ACTION act_Status:
IF TRUE 
AND fbPis.m_CheckByRecipe(stPis:=stPis_TankA, 			req:=E_Piston_Recipe_State.Release)	
//AND fbPis.m_CheckByRecipe(stPis:=stPis_TankA_Pipe, 		req:=E_Piston_Recipe_State.Release)	
AND fbPis.m_CheckByRecipe(stPis:=stPis_TankB, 			req:=E_Piston_Recipe_State.Release)
//AND fbPis.m_CheckByRecipe(stPis:=stPis_TankB_Pipe, 		req:=E_Piston_Recipe_State.Release)
AND fbPis.m_CheckByRecipe(stPis:=stPis_Drain, 			req:=E_Piston_Recipe_State.Release)
AND fbPis.m_CheckByRecipe(stPis:=stPis_CIP, 			req:=E_Piston_Recipe_State.Release)
THEN;
	eStatus:=E_Line_Target.eClose;
ELSIF TRUE 
AND fbPis.m_CheckByRecipe(stPis:=stPis_TankA, 			req:=E_Piston_Recipe_State.Act)		
AND fbPis.m_CheckByRecipe(stPis:=stPis_TankA_Pipe, 		req:=E_Piston_Recipe_State.Release)	
AND fbPis.m_CheckByRecipe(stPis:=stPis_TankB, 			req:=E_Piston_Recipe_State.Release)
//AND fbPis.m_CheckByRecipe(stPis:=stPis_TankB_Pipe, 		req:=E_Piston_Recipe_State.Release)
AND fbPis.m_CheckByRecipe(stPis:=stPis_Drain, 			req:=E_Piston_Recipe_State.Release)
AND fbPis.m_CheckByRecipe(stPis:=stPis_CIP, 			req:=E_Piston_Recipe_State.Release)
THEN;
	eStatus:=E_Line_Target.eTank_A;
ELSIF TRUE 
AND fbPis.m_CheckByRecipe(stPis:=stPis_TankA, 			req:=E_Piston_Recipe_State.Release)		
//AND fbPis.m_CheckByRecipe(stPis:=stPis_TankA_Pipe, 		req:=E_Piston_Recipe_State.Release)	
AND fbPis.m_CheckByRecipe(stPis:=stPis_TankB, 			req:=E_Piston_Recipe_State.Act)
AND fbPis.m_CheckByRecipe(stPis:=stPis_TankB_Pipe, 		req:=E_Piston_Recipe_State.Release)
AND fbPis.m_CheckByRecipe(stPis:=stPis_Drain, 			req:=E_Piston_Recipe_State.Release)
AND fbPis.m_CheckByRecipe(stPis:=stPis_CIP, 			req:=E_Piston_Recipe_State.Release)
THEN;
	eStatus:=E_Line_Target.eTank_B;
ELSIF TRUE 
AND fbPis.m_CheckByRecipe(stPis:=stPis_TankA, 			req:=E_Piston_Recipe_State.Release)		
//AND fbPis.m_CheckByRecipe(stPis:=stPis_TankA_Pipe, 		req:=E_Piston_Recipe_State.Release)	
AND fbPis.m_CheckByRecipe(stPis:=stPis_TankB, 			req:=E_Piston_Recipe_State.Release)
//AND fbPis.m_CheckByRecipe(stPis:=stPis_TankB_Pipe, 		req:=E_Piston_Recipe_State.Release)
AND fbPis.m_CheckByRecipe(stPis:=stPis_Drain, 			req:=E_Piston_Recipe_State.Act)
AND fbPis.m_CheckByRecipe(stPis:=stPis_CIP, 			req:=E_Piston_Recipe_State.Act)
THEN;
	eStatus:=E_Line_Target.eCIP;
ELSIF TRUE 
AND fbPis.m_CheckByRecipe(stPis:=stPis_TankA, 			req:=E_Piston_Recipe_State.Release)		
//AND fbPis.m_CheckByRecipe(stPis:=stPis_TankA_Pipe, 		req:=E_Piston_Recipe_State.Release)	
AND fbPis.m_CheckByRecipe(stPis:=stPis_TankB, 			req:=E_Piston_Recipe_State.Release)
//AND fbPis.m_CheckByRecipe(stPis:=stPis_TankB_Pipe, 		req:=E_Piston_Recipe_State.Release)
AND fbPis.m_CheckByRecipe(stPis:=stPis_Drain, 			req:=E_Piston_Recipe_State.Act)
AND fbPis.m_CheckByRecipe(stPis:=stPis_CIP, 			req:=E_Piston_Recipe_State.Release)
THEN;
	eStatus:=E_Line_Target.eDrain;
ELSE;
	eStatus:=E_Line_Target.eNone;
END_IF
END_ACTION

METHOD m_CheckStatus : BOOL
VAR_INPUT
	eReqStatus		: E_Line_Target;
END_VAR
IF eStatus=eReqStatus 
AND eProcess=E_Line_Target.eNone
AND eReq=E_Line_Target.eNone
AND bReady
AND bDone
AND NOT bRun
THEN;
	m_CheckStatus:=TRUE;
END_IF
END_METHOD

METHOD m_Request_Reset : BOOL
VAR_IN_OUT
	memo: R_TRIG;
END_VAR
memo(CLK:=eReq=0);
IF TRUE 
AND memo.Q
THEN;
	SFCReset:=TRUE;
END_IF
END_METHOD

METHOD m_Run : BOOL
VAR_INPUT
	eReqProc			: E_Line_Target;
END_VAR
IF eProcess=E_Line_Target.eNone THEN;
	eProcess:=eReq:=eReqProc;
	bDone:=FALSE;
	m_Run:=TRUE;
END_IF
END_METHOD

METHOD m_Set_SFCFlags_Reference : BOOL
//Set reference to SFC flags

refSFC.SFCInit REF= SFCInit;
refSFC.SFCReset REF= SFCReset;
refSFC.SFCError REF= SFCError;
refSFC.SFCEnableLimit REF= SFCEnableLimit;
refSFC.SFCErrorStep REF= SFCErrorStep;
refSFC.SFCErrorPOU REF= SFCErrorPOU;
refSFC.SFCQuitError REF= SFCQuitError;
refSFC.SFCPause REF= SFCPause;
refSFC.SFCTrans REF= SFCTrans;
refSFC.SFCCurrentStep REF= SFCCurrentStep;
refSFC.SFCTip REF= SFCTip;
refSFC.SFCTipMode REF= SFCTipMode;

// Cycle handle for SFC
m_SFC_Handle();
END_METHOD

END_FUNCTION_BLOCK

// ---- 00 Library/02 Pump/FB_Pump.TcPOU
FUNCTION_BLOCK FB_Pump
VAR_INPUT
	Pump_ID				: E_Pump_List:=E_Pump_List.eNotSelected;
	PressureSensor_ID	: E_ASense_Name:=E_ASense_Name.eNotSelected;
END_VAR
VAR
	sID: STRING(6);

	stNidec: REFERENCE TO ST_Nidec;
	status_word: WORD;
	control_word: WORD;

	ControlWord: ControlWordStruct;
	StatusWord: StatusWordStruct;


	//request
	modeAuto	:	BOOL	:= TRUE	;//System in automatic
	bRun_Auto	:	BOOL	;
	bRun_Man	:	BOOL	;

	//nRPM_Auto	:	REAL		;//Pump RPM 
	//nRPM_Man	:	REAL		;//Pump RPM 
	//feedback
	nRPM_fdbk	:	INT	;	
	rtManual: R_TRIG;
	ton_Drive_init: TON;
	state_init: (OFF,stage1,stage2,stage3,stage4, Ready);

	bInitiated: BOOL;
	ton_RPM_feedback_lag_monitoring: TON;
	ton_Pressure_feedback_monitoring: TON;
	
	fbPressureSensor: REFERENCE TO FB_AnalogSensor;

END_VAR
VAR_OUTPUT
	DriveReady	:   BOOL;
	bRun		: 	BOOL;
	nRPM		:	REAL		;//Pump RPM 
	
END_VAR
VAR_IN_OUT
	stPump			: ST_Pump	;
	stOperation		: ST_OperationButtons;
END_VAR

stNidec REF= gIO.Nidec[Pump_ID];
sID:=TO_STRING(Pump_ID);
nRPM:=stPump.nRPM;
IF __ISVALIDREF(stNidec) THEN;
	//run
	status_word:=stNidec.StatusWord;
	stNidec.ControlWord:=control_word;
	
	control_word:=m_Map_ControlWord(cwStruct:=ControlWord);
	StatusWord:=m_Map_StatusWord(wordInput:=status_word);
	
	stNidec.targetVelocity:=DINT_TO_INT(TRUNC(stPump.nRPM));	
	nRPM_fdbk:=stNidec.actVelocity;	
	
	m_Nidec_Init();
	
	IF state_init=Ready THEN;
		DriveReady:=TRUE;
		ControlWord.EnableOperation:=bRun;
	ELSE;
		DriveReady:=FALSE;
		//bRun:=bRun_Man:=bRun_Auto:=FALSE;
		ControlWord.EnableOperation:=FALSE;
	END_IF	
	stPump.DriveReady:=DriveReady;
ELSE;
	//RETURN;
END_IF

IF modeAuto THEN;
	//bRun:=bRun_Auto;
	IF bRun_Auto AND m_CheckOper() THEN;
		bRun:=TRUE;
	ELSE;
		bRun:=FALSE;
	END_IF
	stPump.nRPM:=stPump.nRPM_Auto;
ELSE;
	//bRun:=bRun_Man;
	IF bRun_Man AND m_CheckOper() THEN;
		bRun:=TRUE;
	ELSE;
		bRun:=FALSE;
	END_IF	
	stPump.nRPM:=stPump.nRPM_Man;
END_IF

rtManual(CLK:=NOT modeAuto);
IF rtManual.Q THEN;
	bRun:=bRun_Man:=bRun_Auto;
	//stPump.nRPM:=stPump.nRPM_Man:=stPump.nRPM_Auto;
END_IF

IF stPump.nRPM>3000 THEN;
	stPump.nRPM:=3000;
END_IF

stPump.bRun_Man:=bRun_Man;
stPump.bRun_Auto:=bRun_Auto;
stPump.bRun:=bRun;

IF m_Error()<>'' THEN;
	//stOperation.bSetPause:=TRUE;
	//print error
	//fbPrintErrMessageByID(sModuleDescription:='Pump',sActErrorID:='101x000x001');	
END_IF

bInitiated:=TRUE;

METHOD m_Auto : BOOL
VAR_INPUT
	control: LREAL; // RPM
END_VAR

VAR
	RPM: INT;
END_VAR
//ST_Pump.bRun_Auto:=TRUE;
m_Auto:=TRUE;
RPM:=DINT_TO_INT(TRUNC(control));
IF RPM>3000 THEN;
	stPump.nRPM_Auto:=3000;
ELSIF RPM<200 THEN;
	stPump.nRPM_Auto:=200;
ELSE;
	stPump.nRPM_Auto:=RPM;
END_IF

bRun_Auto:=TRUE;
//need to be set up an set point so the pump could keep the needed value in automatic mode
END_METHOD

METHOD INTERNAL m_CheckOper : BOOL
VAR_INPUT
END_VAR

VAR
	sMotorTypeAgrigate_to_check: STRING(2);
END_VAR
sMotorTypeAgrigate_to_check:=TO_STRING(Pump_ID);

IF sMotorTypeAgrigate_to_check='AG' THEN;
	m_CheckOper:=TRUE;
ELSE;
	IF stOperation.iActOperation=E_OperationButtons.ePlayAll THEN;
		m_CheckOper:=TRUE;
	ELSE;
		m_CheckOper:=FALSE;
	END_IF
END_IF
END_METHOD

METHOD m_Error : STRING(11)
VAR_INPUT
	
END_VAR
VAR
	skipTemp: BOOL;
END_VAR
ton_RPM_feedback_lag_monitoring(PT:=T#10S);
IF __ISVALIDREF(stNidec) THEN;
	IF bRun
	AND ABS(stNidec.targetVelocity - nRPM_fdbk) > 10 
	THEN;
		ton_RPM_feedback_lag_monitoring.IN:=TRUE;
	ELSE;
		ton_RPM_feedback_lag_monitoring.IN:=FALSE;
	END_IF	
END_IF

CASE Pump_ID OF
	E_Pump_List.AG3001,
	E_Pump_List.AG3002,
	E_Pump_List.P3001,
	E_Pump_List.P3002:;
		skipTemp:=TRUE;
ELSE;
		skipTemp:=FALSE;
END_CASE


IF bRun AND NOT skipTemp THEN;
	IF NOT DriveReady THEN;
		m_Error:=concat(sID,'x001');
		stOperation.bSetPause:=TRUE;
		RETURN;
	END_IF	

	IF ton_RPM_feedback_lag_monitoring.Q THEN;
		m_Error:=concat(sID,'x002');
		RETURN;
	END_IF
END_IF

IF NOT DriveReady AND NOT skipTemp THEN;
	m_Error:=concat(sID,'x003');
	//stOperation.bSetPause:=TRUE;
	RETURN;
END_IF


IF 	PressureSensor_ID <> E_ASense_Name.eNotSelected THEN;
	fbPressureSensor REF= fbAnalogSensor[PressureSensor_ID];
	IF __ISVALIDREF(fbPressureSensor) THEN;	
		ton_Pressure_feedback_monitoring(PT:=T#30S);
		IF bRun AND ( fbPressureSensor.bHH_Alarm 
					OR fbPressureSensor.bHH_Warning
					OR fbPressureSensor.bLL_Warning 
					OR fbPressureSensor.bLL_Alarm) 
		THEN;
			ton_Pressure_feedback_monitoring.IN:=TRUE;
		ELSE;
			ton_Pressure_feedback_monitoring.IN:=FALSE;
		END_IF	
		
		IF fbPressureSensor.bHH_Alarm AND ton_Pressure_feedback_monitoring.Q THEN;
			m_Error:=concat(sID,'x004');
			stOperation.bSetPause:=TRUE;
			RETURN;
		END_IF
		IF fbPressureSensor.bHH_Warning AND ton_Pressure_feedback_monitoring.Q THEN;
			m_Error:=concat(sID,'x005');
			RETURN;
		END_IF
		IF fbPressureSensor.bLL_Warning AND ton_Pressure_feedback_monitoring.Q THEN;
			m_Error:=concat(sID,'x006');
			RETURN;
		END_IF
		IF fbPressureSensor.bLL_Alarm AND ton_Pressure_feedback_monitoring.Q THEN;
			m_Error:=concat(sID,'x007');
			stOperation.bSetPause:=TRUE;
			RETURN;
		END_IF		
	END_IF	
END_IF

IF NOT modeAuto THEN;
	m_Error:=concat(sID,'x008');
	//stOperation.bSetPause:=TRUE;
	RETURN;
END_IF

m_Error:='';
END_METHOD

METHOD m_Get_Speed : INT
VAR_INPUT
END_VAR
m_Get_Speed:=nRPM_fdbk;
END_METHOD

METHOD m_Map_ControlWord : WORD
VAR_INPUT
	cwStruct : ControlWordStruct;
END_VAR
VAR
    tempWord : WORD;
END_VAR


// Map each bit from the structure to the corresponding bit in the control word
tempWord := 0;
IF cwStruct.SwitchOn THEN
    tempWord := tempWord OR 1; // Bit 0
END_IF
IF cwStruct.EnableVoltage THEN
    tempWord := tempWord OR 2; // Bit 1
END_IF
IF cwStruct.QuickStop THEN
    tempWord := tempWord OR 4; // Bit 2
END_IF
IF cwStruct.EnableOperation THEN
    tempWord := tempWord OR 8; // Bit 3
END_IF
// Reserved bits (4-7) are not set
IF cwStruct.FaultReset THEN
    tempWord := tempWord OR 256; // Bit 8
END_IF
// Reserved bits (9-15) are not set

m_Map_ControlWord := tempWord;
END_METHOD

METHOD m_Map_StatusWord : StatusWordStruct
VAR_INPUT
	wordInput : WORD;
END_VAR
VAR
    swStruct : StatusWordStruct;
END_VAR


// Map each bit from the status word to the corresponding field in the structure
swStruct.ReadyToSwitchOn    := (wordInput AND 1) <> 0;         // Bit 0
swStruct.SwitchedOn         := (wordInput AND 2) <> 0;         // Bit 1
swStruct.OperationEnabled   := (wordInput AND 4) <> 0;         // Bit 2
swStruct.Fault              := (wordInput AND 8) <> 0;         // Bit 3
swStruct.VoltageEnabled     := (wordInput AND 16) <> 0;        // Bit 4
swStruct.QuickStop          := (wordInput AND 32) <> 0;        // Bit 5
swStruct.SwitchOnDisabled   := (wordInput AND 64) <> 0;        // Bit 6
swStruct.Warning            := (wordInput AND 128) <> 0;       // Bit 7
swStruct.Remote             := (wordInput AND 256) <> 0;       // Bit 8
// Reserved bits (9-15) are not set, assuming FALSE
m_Map_StatusWord := swStruct;
END_METHOD

METHOD m_Nidec_Init : BOOL
VAR_INPUT
END_VAR
IF  NOT StatusWord.VoltageEnabled 
OR StatusWord.Fault 
OR (state_init=Ready AND NOT StatusWord.ReadyToSwitchOn )
THEN;
	ControlWord.SwitchOn:=FALSE;
	ControlWord.EnableVoltage:=FALSE;
	ControlWord.QuickStop:=FALSE;
	ControlWord.EnableOperation:=FALSE;
	ton_Drive_init(IN:=FALSE);
	state_init:=OFF;
	RETURN;
END_IF


CASE state_init OF
	OFF:; 
		IF TRUE
		AND StatusWord.VoltageEnabled
		AND StatusWord.QuickStop
		AND StatusWord.SwitchOnDisabled
		THEN;
			ton_Drive_init(IN:=TRUE,PT:=T#2S);
		ELSE;
			ton_Drive_init(IN:=FALSE);RETURN;
		END_IF
		
		IF ton_Drive_init.Q THEN;
			ControlWord.EnableVoltage:=TRUE;
			ControlWord.QuickStop:=TRUE;	
			state_init:=stage1;
			ton_Drive_init(IN:=FALSE);
		END_IF	
		
	stage1:;
		IF TRUE
		AND StatusWord.VoltageEnabled
		AND StatusWord.QuickStop
		AND NOT StatusWord.SwitchOnDisabled
		THEN;
			ton_Drive_init(IN:=TRUE,PT:=T#0.5S);
		ELSE;
			ton_Drive_init(IN:=FALSE);RETURN;
		END_IF
		
		IF ton_Drive_init.Q THEN;
			ControlWord.SwitchOn:=TRUE;
			state_init:=stage2;
			ton_Drive_init(IN:=FALSE);
		END_IF	
		
	stage2:;
		IF TRUE
		AND StatusWord.SwitchedOn
		AND StatusWord.VoltageEnabled
		AND StatusWord.QuickStop
		AND NOT StatusWord.SwitchOnDisabled
		THEN;
			ton_Drive_init(IN:=TRUE,PT:=T#0.5S);
		ELSE;
			ton_Drive_init(IN:=FALSE);RETURN;
		END_IF
		
		IF ton_Drive_init.Q THEN;
			state_init:=Ready;
			ton_Drive_init(IN:=FALSE);
		END_IF	

	
	
END_CASE
END_METHOD

METHOD m_Run : BOOL
VAR_INPUT
	RPM: REAL;
END_VAR
IF NOT bInitiated THEN;
	RETURN;
END_IF
bRun_Auto:=TRUE;
stPump.nRPM_Auto:=RPM;
m_Run:=TRUE;
END_METHOD

METHOD m_Stop : BOOL
VAR_INPUT
END_VAR
bRun_Auto:=FALSE;
bRun_Man:=FALSE;
m_Stop:=TRUE;
END_METHOD

END_FUNCTION_BLOCK

// ---- 00 Library/02 Pump/02.1 Dosing Pump/FB_DosingPump.TcPOU
FUNCTION_BLOCK FB_DosingPump EXTENDS FB_SFC_Cycle
VAR_INPUT
END_VAR
VAR_OUTPUT
	valve_A			: BOOL;
	valve_B			: BOOL;
END_VAR
VAR

	action_Time		: TIME:=T#0.5S;
	startDelay		: TIME:=T#0S;
	
	reqTiks			: DINT:=5;
	actTiks			: DINT:=5;
	
	fStageVolume	: REAL:=65; 	// CC/stage
	fReqVolume		: REAL:=500.0; 	// CC
	fActVolume		: REAL; 		// CC


END_VAR

VAR PERSISTENT
	
END_VAR

act_GetReference();

act_Oper();

reqTiks:=TRUNC(fReqVolume/fStageVolume);
fActVolume:=(actTiks*fStageVolume);

ACTION _acheck_Count_active:
bStepDone:=FALSE;
IF actTiks>=reqTiks THEN;
	bStepDone:=TRUE;
END_IF
END_ACTION

ACTION _acheck_Count_entry:
actTiks:=actTiks+1;
END_ACTION

ACTION _aDone_entry:
bRun:=FALSE;
bDone:=TRUE;
END_ACTION

ACTION _aInit_act_Oper_active:
SFCReset:=FALSE;
END_ACTION

ACTION _aInit_act_Oper_exit:
valve_A:=valve_B:=bRun:=bDone:=FALSE;
END_ACTION

ACTION _aReady_exit:
actTiks:=0;
END_ACTION

ACTION _astage_A_entry:
valve_A:=TRUE;
END_ACTION

ACTION _astage_A_exit:
valve_A:=FALSE;
END_ACTION

ACTION _astage_B_entry:
valve_B:=TRUE;
END_ACTION

ACTION _astage_B_exit:
valve_B:=FALSE;
END_ACTION

ACTION act_GetReference:
m_Set_SFCFlags_Reference();
END_ACTION

ACTION act_Oper:
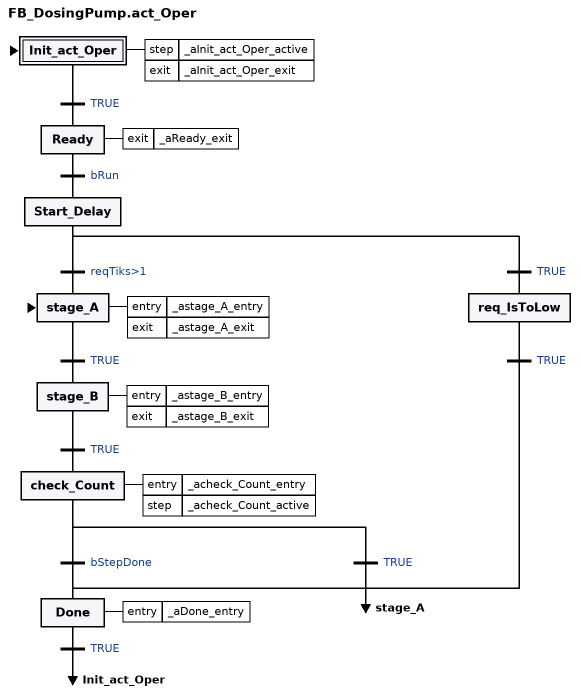
INITIAL_STEP Init_act_Oper:
    _aInit_act_Oper_active(N);  // step action
    _aInit_act_Oper_exit(P0);  // exit action
END_STEP
TRANSITION FROM Init_act_Oper TO Ready
    := TRUE;
END_TRANSITION
STEP Ready:
    _aReady_exit(P0);  // exit action
END_STEP
TRANSITION FROM Ready TO Start_Delay
    := bRun;
END_TRANSITION
STEP Start_Delay:  // min time startDelay
END_STEP
TRANSITION FROM Start_Delay TO stage_A
    := reqTiks>1;
END_TRANSITION
STEP stage_A:  // min time action_Time
    _astage_A_entry(P1);  // entry action
    _astage_A_exit(P0);  // exit action
END_STEP
TRANSITION FROM stage_A TO stage_B
    := TRUE;
END_TRANSITION
STEP stage_B:  // min time action_Time
    _astage_B_entry(P1);  // entry action
    _astage_B_exit(P0);  // exit action
END_STEP
TRANSITION FROM stage_B TO check_Count
    := TRUE;
END_TRANSITION
STEP check_Count:
    _acheck_Count_entry(P1);  // entry action
    _acheck_Count_active(N);  // step action
END_STEP
TRANSITION FROM check_Count TO Done
    := bStepDone;
END_TRANSITION
TRANSITION FROM check_Count TO stage_A
    := TRUE;
END_TRANSITION
TRANSITION FROM Start_Delay TO req_IsToLow
    := TRUE;
END_TRANSITION
STEP req_IsToLow:
END_STEP
TRANSITION FROM req_IsToLow TO Done
    := TRUE;
END_TRANSITION
STEP Done:
    _aDone_entry(P1);  // entry action
END_STEP
TRANSITION FROM Done TO Init_act_Oper
    := TRUE;
END_TRANSITION
// branch label Branch0_act_Oper
// branch label Branch1_act_Oper
END_ACTION

METHOD m_RunVolume : BOOL
VAR_INPUT
	Volume	:REAL;
END_VAR
fReqVolume:=Volume;
mRun();
IF rtDone.Q THEN;
	m_RunVolume:=TRUE;	
END_IF
END_METHOD

METHOD m_Set_SFCFlags_Reference : BOOL
//Set reference to SFC flags

refSFC.SFCInit REF= SFCInit;
refSFC.SFCReset REF= SFCReset;
refSFC.SFCError REF= SFCError;
refSFC.SFCEnableLimit REF= SFCEnableLimit;
refSFC.SFCErrorStep REF= SFCErrorStep;
refSFC.SFCErrorPOU REF= SFCErrorPOU;
refSFC.SFCQuitError REF= SFCQuitError;
refSFC.SFCPause REF= SFCPause;
refSFC.SFCTrans REF= SFCTrans;
refSFC.SFCCurrentStep REF= SFCCurrentStep;
refSFC.SFCTip REF= SFCTip;
refSFC.SFCTipMode REF= SFCTipMode;

// Cycle handle for SFC
m_SFC_Handle();
END_METHOD

METHOD m_Stop : BOOL
VAR_INPUT
END_VAR
SFCReset:=TRUE;
END_METHOD

END_FUNCTION_BLOCK

// ---- 00 Library/HeatExchenger/FB_HeatExchanger.TcPOU
FUNCTION_BLOCK FB_HeatExchanger
VAR_IN_OUT
	stHeatExchanger	:	ST_HeatExchanger	;
END_VAR
VAR_INPUT
	nValveID		:	E_Pis_Name 	;	
	nAnalogValveID	:	E_Pis_Name 	;

	nProcCntrlID	:	E_ProcessControl_Name	;
END_VAR
VAR_OUTPUT
	nAlagonValveCntrOut	:	INT	;//output for analog valve opening
END_VAR
VAR
	stPis			:	REFERENCE TO ST_Piston;
	stPisAnalog		:	REFERENCE TO ST_Piston;
	
	stProcessControl		:	REFERENCE TO ST_ProcessControl	;
	fbProcessControl		: 	REFERENCE TO FB_ProcessControl	;
END_VAR

act_GetReference();
//act_AnalogOutScaling();

stProcessControl.fCtrlOutput_Min:=0;
stProcessControl.fCtrlOutput_Max:=100;
stProcessControl.fCtrlOutput_Manual;
stProcessControl.rValue_Min_To_ReleaseControl:=15; //Degrees

IF stHeatExchanger.bManual THEN;
	fbProcessControl.mRun_PID(Set_Point:=stProcessControl.fCtrlOutput_Manual , controlManual:=TRUE);
	//nAlagonValveCntrOut:=mCMD_to_Analog(fControl:=stHeatExchanger.fManualControl);
ELSE;
	IF stProcessControl.bActiveCntr AND NOT stPis.st_Open THEN
		stPis.req_Open:=TRUE;
	ELSIF NOT stProcessControl.bActiveCntr AND NOT stPis.st_Close THEN
		stPis.req_Close:=TRUE;
	END_IF
	//nAlagonValveCntrOut:=mCMD_to_Analog(fControl:=stProcessControl.fCtrlOutput);	
END_IF
nAlagonValveCntrOut:=mCMD_to_Analog(fControl:=stProcessControl.fCtrlOutput);
IF nAlagonValveCntrOut=0 AND NOT stPisAnalog.st_Close THEN;
	stPisAnalog.req_Close:=TRUE;
ELSIF nAlagonValveCntrOut<>0 AND NOT stPisAnalog.st_Open THEN;
	stPisAnalog.req_Open:=TRUE;
END_IF

ACTION act_AnalogOutScaling:
IF (stHeatExchanger.cntrlVal_Max-stHeatExchanger.cntrlVal_Min)<>0 THEN
	nAlagonValveCntrOut:=DINT_TO_INT((TRUNC((stProcessControl.fCtrlOutput*
		(stHeatExchanger.outVal_Max-stHeatExchanger.outVal_Min)/(stHeatExchanger.cntrlVal_Max-stHeatExchanger.cntrlVal_Min))+
		stHeatExchanger.outOffset)));
END_IF
END_ACTION

ACTION act_GetReference:
//On-Off walve structure
stPis REF= g_Piston.stPis[nValveID];
stPisAnalog REF= g_Piston.stPis[nAnalogValveID];

stProcessControl REF=g_ProcControl.arr_stProcCntrl[nProcCntrlID];
fbProcessControl REF=g_ProcControl.arr_fbProcCntrl[nProcCntrlID];
END_ACTION

METHOD m_Auto : BOOL
VAR_INPUT
END_VAR
END_METHOD

METHOD m_Run : BOOL
VAR_INPUT
END_VAR
END_METHOD

METHOD m_Stop : BOOL
VAR_INPUT
END_VAR
END_METHOD

METHOD mCMD_to_Analog : INT
VAR_INPUT
	fControl: LREAL;
END_VAR
IF (stHeatExchanger.cntrlVal_Max-stHeatExchanger.cntrlVal_Min)<>0 THEN
	mCMD_to_Analog:=DINT_TO_INT((TRUNC((fControl*
		(stHeatExchanger.outVal_Max-stHeatExchanger.outVal_Min)/(stHeatExchanger.cntrlVal_Max-stHeatExchanger.cntrlVal_Min))+
		stHeatExchanger.outOffset)));
ELSE;
	mCMD_to_Analog:=0;
END_IF

//nAlagonValveCntrOut
END_METHOD

END_FUNCTION_BLOCK

// ---- 03 Project/23 CIP/FB_CIP_ClientTank.TcPOU
FUNCTION_BLOCK FB_CIP_ClientTank EXTENDS FB_SFC_Cycle IMPLEMENTS ITF_FB_SFC_Cycle
VAR_INPUT	
	valTank_A				: E_Pis_Name;
	valTank_A_Sprinkler		: E_Pis_Name;
	valTank_A_Main			: E_Pis_Name;
	valTank_B				: E_Pis_Name;
	valTank_B_Sprinkler		: E_Pis_Name;	
	valTank_B_Main			: E_Pis_Name;	
	valDrain				: E_Pis_Name;
END_VAR
VAR_OUTPUT
END_VAR
VAR

	eReq				: E_CIP_ClientTank;
	eProcess			: E_CIP_ClientTank;
	eStatus				: E_CIP_ClientTank;
	
	fbPis					: FB_Piston;
	stPis_Tank_A			: REFERENCE TO ST_Piston;
	stPis_Tank_A_Sprinkler	: REFERENCE TO ST_Piston;
	stPis_Tank_A_Main		: REFERENCE TO ST_Piston;
	stPis_Tank_B			: REFERENCE TO ST_Piston;
	stPis_Tank_B_Sprinkler	: REFERENCE TO ST_Piston;
	stPis_Tank_B_Main		: REFERENCE TO ST_Piston;
	stPis_Drain				: REFERENCE TO ST_Piston;

	tonDrainTime: TON;
	rt_Req_Reset: R_TRIG;
END_VAR
VAR_IN_OUT


END_VAR

act_GetReference();

act_Oper();
IF NOT Init.x THEN;
	act_Status();
END_IF

tonDrainTime(PT:=T#1M, IN:=eStatus=E_CIP_ClientTank.eDrain);
IF tonDrainTime.Q 
AND eReq=E_CIP_ClientTank.eNone
AND eProcess=E_CIP_ClientTank.eNone
THEN;
	eReq:=E_CIP_ClientTank.eClose;
END_IF

m_Request_Reset(memo:=rt_Req_Reset);

ACTION _aClose_active:
bStepDone:=FALSE;
IF TRUE 
AND eStatus=E_CIP_ClientTank.eClose
THEN;
	bStepDone:=TRUE;
END_IF
END_ACTION

ACTION _aClose_entry:
fbPis.m_SetByRecipe(stPis:=stPis_Tank_A, 				req:=E_Piston_Recipe_State.Release);
fbPis.m_SetByRecipe(stPis:=stPis_Tank_A_Sprinkler, 		req:=E_Piston_Recipe_State.Release);
fbPis.m_SetByRecipe(stPis:=stPis_Tank_A_Main, 			req:=E_Piston_Recipe_State.Release);
fbPis.m_SetByRecipe(stPis:=stPis_Tank_B, 				req:=E_Piston_Recipe_State.Release);
fbPis.m_SetByRecipe(stPis:=stPis_Tank_B_Sprinkler, 		req:=E_Piston_Recipe_State.Release);
fbPis.m_SetByRecipe(stPis:=stPis_Tank_B_Main, 			req:=E_Piston_Recipe_State.Release);
fbPis.m_SetByRecipe(stPis:=stPis_Drain, 				req:=E_Piston_Recipe_State.Release);
END_ACTION

ACTION _aDone_entry:
eProcess:=E_CIP_ClientTank.eNone;
eReq:=E_CIP_ClientTank.eNone;
bRun:=FALSE;
bDone:=TRUE;
END_ACTION

ACTION _aDrain_active:
bStepDone:=FALSE;
IF TRUE 
AND eStatus=E_CIP_ClientTank.eDrain
THEN;
	bStepDone:=TRUE;
END_IF
END_ACTION

ACTION _aDrain_entry:
fbPis.m_SetByRecipe(stPis:=stPis_Tank_A, 				req:=E_Piston_Recipe_State.Release);
fbPis.m_SetByRecipe(stPis:=stPis_Tank_A_Sprinkler, 		req:=E_Piston_Recipe_State.Release);
fbPis.m_SetByRecipe(stPis:=stPis_Tank_A_Main, 			req:=E_Piston_Recipe_State.Release);
fbPis.m_SetByRecipe(stPis:=stPis_Tank_B, 				req:=E_Piston_Recipe_State.Release);
fbPis.m_SetByRecipe(stPis:=stPis_Tank_B_Sprinkler, 		req:=E_Piston_Recipe_State.Release);
fbPis.m_SetByRecipe(stPis:=stPis_Tank_B_Main, 			req:=E_Piston_Recipe_State.Release);
fbPis.m_SetByRecipe(stPis:=stPis_Drain, 				req:=E_Piston_Recipe_State.Act);
END_ACTION

ACTION _aInit_active:
SFCReset:=FALSE;
END_ACTION

ACTION _aInit_exit:
eProcess:=E_CIP_ClientTank.eNone;
eReq:=E_CIP_ClientTank.eNone;
END_ACTION

ACTION _aReady_active:


CASE eReq OF
	E_CIP_ClientTank.eClose:;
			IF TRUE THEN;
				eProcess:=E_CIP_ClientTank.eClose;
			END_IF

	E_CIP_ClientTank.eTank_A:;
			IF TRUE THEN;
				eProcess:=E_CIP_ClientTank.eTank_A;
			END_IF	
			
	E_CIP_ClientTank.eTank_A_Sprinkler:;
			IF TRUE THEN;
				eProcess:=E_CIP_ClientTank.eTank_A_Sprinkler;
			END_IF
			
	E_CIP_ClientTank.eTank_B:;
			IF TRUE THEN;
				eProcess:=E_CIP_ClientTank.eTank_B;
			END_IF	
	
	E_CIP_ClientTank.eTank_B_Sprinkler:;
			IF TRUE THEN;
				eProcess:=E_CIP_ClientTank.eTank_B_Sprinkler;
			END_IF	

	E_CIP_ClientTank.eDrain:;
			IF TRUE THEN;
				eProcess:=E_CIP_ClientTank.eDrain;
			END_IF	
	

END_CASE
END_ACTION

ACTION _aReady_exit:
bRun:=TRUE;
bDone:=FALSE;
END_ACTION

ACTION _aTank_A_active:
bStepDone:=FALSE;
IF TRUE 
AND eStatus=E_CIP_ClientTank.eTank_A
THEN;
	bStepDone:=TRUE;
END_IF
END_ACTION

ACTION _aTank_A_entry:
fbPis.m_SetByRecipe(stPis:=stPis_Tank_A, 				req:=E_Piston_Recipe_State.Act);
fbPis.m_SetByRecipe(stPis:=stPis_Tank_A_Sprinkler, 		req:=E_Piston_Recipe_State.Release);
fbPis.m_SetByRecipe(stPis:=stPis_Tank_A_Main, 			req:=E_Piston_Recipe_State.Release);
fbPis.m_SetByRecipe(stPis:=stPis_Tank_B, 				req:=E_Piston_Recipe_State.Release);
fbPis.m_SetByRecipe(stPis:=stPis_Tank_B_Sprinkler, 		req:=E_Piston_Recipe_State.Release);
fbPis.m_SetByRecipe(stPis:=stPis_Tank_B_Main, 			req:=E_Piston_Recipe_State.Release);
fbPis.m_SetByRecipe(stPis:=stPis_Drain, 				req:=E_Piston_Recipe_State.Release);
END_ACTION

ACTION _aTank_A_Sprinkler_active:
bStepDone:=FALSE;
IF TRUE 
AND eStatus=E_CIP_ClientTank.eTank_A_Sprinkler
THEN;
	bStepDone:=TRUE;
END_IF
END_ACTION

ACTION _aTank_A_Sprinkler_entry:
fbPis.m_SetByRecipe(stPis:=stPis_Tank_A, 				req:=E_Piston_Recipe_State.Act);
fbPis.m_SetByRecipe(stPis:=stPis_Tank_A_Sprinkler, 		req:=E_Piston_Recipe_State.Act);
fbPis.m_SetByRecipe(stPis:=stPis_Tank_A_Main, 			req:=E_Piston_Recipe_State.Act);
fbPis.m_SetByRecipe(stPis:=stPis_Tank_B, 				req:=E_Piston_Recipe_State.Release);
fbPis.m_SetByRecipe(stPis:=stPis_Tank_B_Sprinkler, 		req:=E_Piston_Recipe_State.Release);
fbPis.m_SetByRecipe(stPis:=stPis_Tank_B_Main, 			req:=E_Piston_Recipe_State.Release);
fbPis.m_SetByRecipe(stPis:=stPis_Drain, 				req:=E_Piston_Recipe_State.Release);
END_ACTION

ACTION _aTank_B_active:
bStepDone:=FALSE;
IF TRUE 
AND eStatus=E_CIP_ClientTank.eTank_B
THEN;
	bStepDone:=TRUE;
END_IF
END_ACTION

ACTION _aTank_B_entry:
fbPis.m_SetByRecipe(stPis:=stPis_Tank_A, 				req:=E_Piston_Recipe_State.Release);
fbPis.m_SetByRecipe(stPis:=stPis_Tank_A_Sprinkler, 		req:=E_Piston_Recipe_State.Release);
fbPis.m_SetByRecipe(stPis:=stPis_Tank_A_Main, 			req:=E_Piston_Recipe_State.Release);
fbPis.m_SetByRecipe(stPis:=stPis_Tank_B, 				req:=E_Piston_Recipe_State.Act);
fbPis.m_SetByRecipe(stPis:=stPis_Tank_B_Sprinkler, 		req:=E_Piston_Recipe_State.Release);
fbPis.m_SetByRecipe(stPis:=stPis_Tank_B_Main, 			req:=E_Piston_Recipe_State.Release);
fbPis.m_SetByRecipe(stPis:=stPis_Drain, 				req:=E_Piston_Recipe_State.Release);
END_ACTION

ACTION _aTank_B_Sprinkler_active:
bStepDone:=FALSE;
IF TRUE 
AND eStatus=E_CIP_ClientTank.eTank_B_Sprinkler
THEN;
	bStepDone:=TRUE;
END_IF
END_ACTION

ACTION _aTank_B_Sprinkler_entry:
fbPis.m_SetByRecipe(stPis:=stPis_Tank_A, 				req:=E_Piston_Recipe_State.Release);
fbPis.m_SetByRecipe(stPis:=stPis_Tank_A_Sprinkler, 		req:=E_Piston_Recipe_State.Release);
fbPis.m_SetByRecipe(stPis:=stPis_Tank_A_Main, 			req:=E_Piston_Recipe_State.Release);
fbPis.m_SetByRecipe(stPis:=stPis_Tank_B, 				req:=E_Piston_Recipe_State.Act);
fbPis.m_SetByRecipe(stPis:=stPis_Tank_B_Sprinkler, 		req:=E_Piston_Recipe_State.Act);
fbPis.m_SetByRecipe(stPis:=stPis_Tank_B_Main, 			req:=E_Piston_Recipe_State.Act);
fbPis.m_SetByRecipe(stPis:=stPis_Drain, 				req:=E_Piston_Recipe_State.Release);
END_ACTION

ACTION act_GetReference:
m_Set_SFCFlags_Reference();
	
stPis_Tank_A				REF= g_Piston.stPis[valTank_A];
stPis_Tank_A_Sprinkler		REF= g_Piston.stPis[valTank_A_Sprinkler];
stPis_Tank_A_Main			REF= g_Piston.stPis[valTank_A_Main];
stPis_Tank_B				REF= g_Piston.stPis[valTank_B];
stPis_Tank_B_Sprinkler		REF= g_Piston.stPis[valTank_B_Sprinkler];
stPis_Tank_B_Main			REF= g_Piston.stPis[valTank_B_Main];
stPis_Drain					REF= g_Piston.stPis[valDrain];
END_ACTION

ACTION act_Oper:
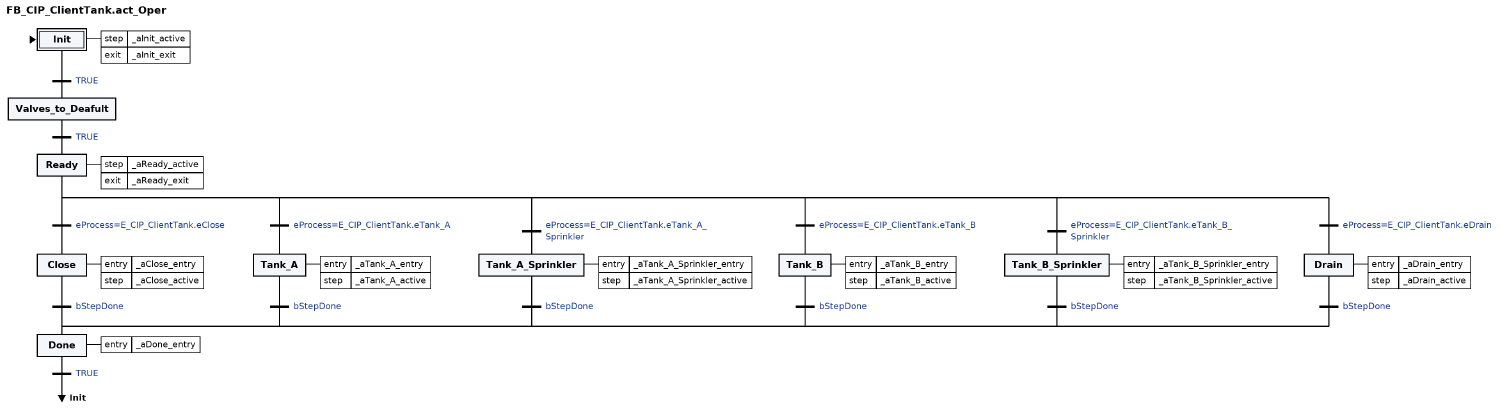
INITIAL_STEP Init:  // min time T#0.5s
    _aInit_active(N);  // step action
    _aInit_exit(P0);  // exit action
END_STEP
TRANSITION FROM Init TO Valves_to_Deafult
    := TRUE;
END_TRANSITION
STEP Valves_to_Deafult:
END_STEP
TRANSITION FROM Valves_to_Deafult TO Ready
    := TRUE;
END_TRANSITION
STEP Ready:
    _aReady_active(N);  // step action
    _aReady_exit(P0);  // exit action
END_STEP
TRANSITION FROM Ready TO Close
    := eProcess=E_CIP_ClientTank.eClose;
END_TRANSITION
STEP Close:
    _aClose_entry(P1);  // entry action
    _aClose_active(N);  // step action
END_STEP
TRANSITION FROM Close TO Done
    := bStepDone;
END_TRANSITION
TRANSITION FROM Ready TO Tank_A
    := eProcess=E_CIP_ClientTank.eTank_A;
END_TRANSITION
STEP Tank_A:
    _aTank_A_entry(P1);  // entry action
    _aTank_A_active(N);  // step action
END_STEP
TRANSITION FROM Tank_A TO Done
    := bStepDone;
END_TRANSITION
TRANSITION FROM Ready TO Tank_A_Sprinkler
    := eProcess=E_CIP_ClientTank.eTank_A_Sprinkler;
END_TRANSITION
STEP Tank_A_Sprinkler:
    _aTank_A_Sprinkler_entry(P1);  // entry action
    _aTank_A_Sprinkler_active(N);  // step action
END_STEP
TRANSITION FROM Tank_A_Sprinkler TO Done
    := bStepDone;
END_TRANSITION
TRANSITION FROM Ready TO Tank_B
    := eProcess=E_CIP_ClientTank.eTank_B;
END_TRANSITION
STEP Tank_B:
    _aTank_B_entry(P1);  // entry action
    _aTank_B_active(N);  // step action
END_STEP
TRANSITION FROM Tank_B TO Done
    := bStepDone;
END_TRANSITION
TRANSITION FROM Ready TO Tank_B_Sprinkler
    := eProcess=E_CIP_ClientTank.eTank_B_Sprinkler;
END_TRANSITION
STEP Tank_B_Sprinkler:
    _aTank_B_Sprinkler_entry(P1);  // entry action
    _aTank_B_Sprinkler_active(N);  // step action
END_STEP
TRANSITION FROM Tank_B_Sprinkler TO Done
    := bStepDone;
END_TRANSITION
TRANSITION FROM Ready TO Drain
    := eProcess=E_CIP_ClientTank.eDrain;
END_TRANSITION
STEP Drain:
    _aDrain_entry(P1);  // entry action
    _aDrain_active(N);  // step action
END_STEP
TRANSITION FROM Drain TO Done
    := bStepDone;
END_TRANSITION
STEP Done:  // min time T#0.2s
    _aDone_entry(P1);  // entry action
END_STEP
TRANSITION FROM Done TO Init
    := TRUE;
END_TRANSITION
// branch label Branch2_act_Oper
END_ACTION

ACTION act_Status:
IF bReady AND bDone OR TRUE THEN;
	IF TRUE 
	AND fbPis.m_CheckByRecipe(stPis:=stPis_Tank_A, 				req:=E_Piston_Recipe_State.Release)
	AND fbPis.m_CheckByRecipe(stPis:=stPis_Tank_A_Sprinkler, 	req:=E_Piston_Recipe_State.Release)
	AND fbPis.m_CheckByRecipe(stPis:=stPis_Tank_A_Main, 		req:=E_Piston_Recipe_State.Release)
	AND fbPis.m_CheckByRecipe(stPis:=stPis_Tank_B, 				req:=E_Piston_Recipe_State.Release)
	AND fbPis.m_CheckByRecipe(stPis:=stPis_Tank_B_Sprinkler, 	req:=E_Piston_Recipe_State.Release)
	AND fbPis.m_CheckByRecipe(stPis:=stPis_Tank_B_Main, 		req:=E_Piston_Recipe_State.Release)
	AND fbPis.m_CheckByRecipe(stPis:=stPis_Drain, 				req:=E_Piston_Recipe_State.Release)
	THEN;
		eStatus:=E_CIP_ClientTank.eClose;
		
	ELSIF TRUE 
	AND fbPis.m_CheckByRecipe(stPis:=stPis_Tank_A, 				req:=E_Piston_Recipe_State.Act)
	AND fbPis.m_CheckByRecipe(stPis:=stPis_Tank_A_Sprinkler, 	req:=E_Piston_Recipe_State.Release)
	AND fbPis.m_CheckByRecipe(stPis:=stPis_Tank_A_Main, 		req:=E_Piston_Recipe_State.Release)
	AND fbPis.m_CheckByRecipe(stPis:=stPis_Tank_B, 				req:=E_Piston_Recipe_State.Release)
	AND fbPis.m_CheckByRecipe(stPis:=stPis_Tank_B_Sprinkler, 	req:=E_Piston_Recipe_State.Release)
	AND fbPis.m_CheckByRecipe(stPis:=stPis_Tank_B_Main, 		req:=E_Piston_Recipe_State.Release)
	AND fbPis.m_CheckByRecipe(stPis:=stPis_Drain, 				req:=E_Piston_Recipe_State.Release)
	THEN;
		eStatus:=E_CIP_ClientTank.eTank_A;
	
	ELSIF TRUE 
	AND fbPis.m_CheckByRecipe(stPis:=stPis_Tank_A, 				req:=E_Piston_Recipe_State.Act)
	AND fbPis.m_CheckByRecipe(stPis:=stPis_Tank_A_Sprinkler, 	req:=E_Piston_Recipe_State.Act)
	AND fbPis.m_CheckByRecipe(stPis:=stPis_Tank_A_Main, 		req:=E_Piston_Recipe_State.Act)
	AND fbPis.m_CheckByRecipe(stPis:=stPis_Tank_B, 				req:=E_Piston_Recipe_State.Release)
	AND fbPis.m_CheckByRecipe(stPis:=stPis_Tank_B_Sprinkler, 	req:=E_Piston_Recipe_State.Release)
	AND fbPis.m_CheckByRecipe(stPis:=stPis_Tank_B_Main, 		req:=E_Piston_Recipe_State.Release)
	AND fbPis.m_CheckByRecipe(stPis:=stPis_Drain, 				req:=E_Piston_Recipe_State.Release)
	THEN;
		eStatus:=E_CIP_ClientTank.eTank_A_Sprinkler;
		
	ELSIF TRUE 
	AND fbPis.m_CheckByRecipe(stPis:=stPis_Tank_A, 				req:=E_Piston_Recipe_State.Release)
	AND fbPis.m_CheckByRecipe(stPis:=stPis_Tank_A_Sprinkler, 	req:=E_Piston_Recipe_State.Release)
	AND fbPis.m_CheckByRecipe(stPis:=stPis_Tank_A_Main, 		req:=E_Piston_Recipe_State.Release)
	AND fbPis.m_CheckByRecipe(stPis:=stPis_Tank_B, 				req:=E_Piston_Recipe_State.Act)
	AND fbPis.m_CheckByRecipe(stPis:=stPis_Tank_B_Sprinkler, 	req:=E_Piston_Recipe_State.Release)
	AND fbPis.m_CheckByRecipe(stPis:=stPis_Tank_B_Main, 		req:=E_Piston_Recipe_State.Release)
	AND fbPis.m_CheckByRecipe(stPis:=stPis_Drain, 				req:=E_Piston_Recipe_State.Release)
	THEN;
		eStatus:=E_CIP_ClientTank.eTank_B;	
		
	ELSIF TRUE 
	AND fbPis.m_CheckByRecipe(stPis:=stPis_Tank_A, 				req:=E_Piston_Recipe_State.Release)
	AND fbPis.m_CheckByRecipe(stPis:=stPis_Tank_A_Sprinkler, 	req:=E_Piston_Recipe_State.Release)
	AND fbPis.m_CheckByRecipe(stPis:=stPis_Tank_A_Main, 		req:=E_Piston_Recipe_State.Release)
	AND fbPis.m_CheckByRecipe(stPis:=stPis_Tank_B, 				req:=E_Piston_Recipe_State.Act)
	AND fbPis.m_CheckByRecipe(stPis:=stPis_Tank_B_Sprinkler, 	req:=E_Piston_Recipe_State.Act)
	AND fbPis.m_CheckByRecipe(stPis:=stPis_Tank_B_Main, 		req:=E_Piston_Recipe_State.Act)
	AND fbPis.m_CheckByRecipe(stPis:=stPis_Drain, 				req:=E_Piston_Recipe_State.Release)
	THEN;
		eStatus:=E_CIP_ClientTank.eTank_B_Sprinkler;
		
	ELSIF TRUE 	
	AND fbPis.m_CheckByRecipe(stPis:=stPis_Tank_A, 				req:=E_Piston_Recipe_State.Release)
	AND fbPis.m_CheckByRecipe(stPis:=stPis_Tank_A_Sprinkler, 	req:=E_Piston_Recipe_State.Release)
	AND fbPis.m_CheckByRecipe(stPis:=stPis_Tank_A_Main, 		req:=E_Piston_Recipe_State.Release)
	AND fbPis.m_CheckByRecipe(stPis:=stPis_Tank_B, 				req:=E_Piston_Recipe_State.Release)
	AND fbPis.m_CheckByRecipe(stPis:=stPis_Tank_B_Sprinkler, 	req:=E_Piston_Recipe_State.Release)
	AND fbPis.m_CheckByRecipe(stPis:=stPis_Tank_B_Main, 		req:=E_Piston_Recipe_State.Release)
	AND fbPis.m_CheckByRecipe(stPis:=stPis_Drain, 				req:=E_Piston_Recipe_State.Act)
	THEN;
		eStatus:=E_CIP_ClientTank.eDrain;
		
	ELSE;
		eStatus:=E_CIP_ClientTank.eNone;
	END_IF
ELSE;
	eStatus:=E_CIP_ClientTank.eNone;
END_IF
END_ACTION

METHOD m_CheckStatus : BOOL
VAR_INPUT
	eReqStatus		: E_CIP_ClientTank;
END_VAR
IF eStatus=eReqStatus 
AND eProcess=E_CIP_ClientTank.eNone
AND eReq=E_CIP_ClientTank.eNone
AND bReady
AND bDone
AND NOT bRun
THEN;
	m_CheckStatus:=TRUE;
END_IF
END_METHOD

METHOD m_Request_Reset : BOOL
VAR_IN_OUT
	memo: R_TRIG;
END_VAR
memo(CLK:=eReq=0);
IF TRUE 
AND memo.Q
THEN;
	SFCReset:=TRUE;
END_IF
END_METHOD

METHOD m_Run : BOOL
VAR_INPUT
	eReqProc			: E_CIP_ClientTank;
END_VAR
IF eProcess=E_CIP_ClientTank.eNone THEN;
	eProcess:=eReq:=eReqProc;
	bDone:=FALSE;
	m_Run:=TRUE;
END_IF
END_METHOD

METHOD m_Set_SFCFlags_Reference : BOOL
//Set reference to SFC flags

refSFC.SFCInit REF= SFCInit;
refSFC.SFCReset REF= SFCReset;
refSFC.SFCError REF= SFCError;
refSFC.SFCEnableLimit REF= SFCEnableLimit;
refSFC.SFCErrorStep REF= SFCErrorStep;
refSFC.SFCErrorPOU REF= SFCErrorPOU;
refSFC.SFCQuitError REF= SFCQuitError;
refSFC.SFCPause REF= SFCPause;
refSFC.SFCTrans REF= SFCTrans;
refSFC.SFCCurrentStep REF= SFCCurrentStep;
refSFC.SFCTip REF= SFCTip;
refSFC.SFCTipMode REF= SFCTipMode;

// Cycle handle for SFC
m_SFC_Handle();
END_METHOD

END_FUNCTION_BLOCK

// ---- 03 Project/12 TriBlender/FB_TriBlender_Select.TcPOU
FUNCTION_BLOCK FB_TriBlender_Select EXTENDS FB_SFC_Cycle IMPLEMENTS ITF_FB_SFC_Cycle
VAR_INPUT
	valInSelect		: E_Pis_Name;
	valInMarinade	: E_Pis_Name;
	valInColor		: E_Pis_Name;
	valOutSelect	: E_Pis_Name;	
	valOutMarinade	: E_Pis_Name;
	valOutColor		: E_Pis_Name;
	valDrain		: E_Pis_Name;
	
END_VAR
VAR_OUTPUT
END_VAR
VAR
	//refElement		: REFERENCE TO FB_Element;
	//refState_Long		: REFERENCE TO E_Element_State_Long;
	eReq				: E_TriBlenderSelect;
	eProcess			: E_TriBlenderSelect;
	eStatus				: E_TriBlenderSelect;
	
	fbPis				: FB_Piston;
	stPis_InSelect		: REFERENCE TO ST_Piston;
	stPis_InMarinade	: REFERENCE TO ST_Piston;
	stPis_InColor		: REFERENCE TO ST_Piston;
	stPis_OutSelect		: REFERENCE TO ST_Piston;
	stPis_OutMarinade	: REFERENCE TO ST_Piston;
	stPis_OutColor		: REFERENCE TO ST_Piston;
	stPis_Drain			: REFERENCE TO ST_Piston;

	tonDrainTime: TON;
	rt_Req_Reset: R_TRIG;
	//bRun: BOOL;
	//bDone: BOOL;
	SFCReset: BOOL;
	//bStepDone: BOOL;
END_VAR
VAR_IN_OUT


END_VAR

act_GetReference();

act_Oper();
IF NOT Init.x THEN;
	act_Status();
END_IF

tonDrainTime(PT:=T#1M, IN:=eStatus=E_TriBlenderSelect.eDrain);
IF tonDrainTime.Q 
AND eReq=E_TriBlenderSelect.eNone
AND eProcess=E_TriBlenderSelect.eNone
THEN;
	eReq:=E_TriBlenderSelect.eMarinade;
END_IF

m_Request_Reset(memo:=rt_Req_Reset);//

ACTION _aColor_1_active:
bStepDone:=FALSE;
IF TRUE 
AND eStatus=E_TriBlenderSelect.eColor
THEN;
	bStepDone:=TRUE;
END_IF
END_ACTION

ACTION _aColor_1_entry:
fbPis.m_SetByRecipe(stPis:=stPis_InSelect, 			req:=E_Piston_Recipe_State.Act);
fbPis.m_SetByRecipe(stPis:=stPis_InMarinade, 		req:=E_Piston_Recipe_State.Release);
fbPis.m_SetByRecipe(stPis:=stPis_InColor, 			req:=E_Piston_Recipe_State.Release);
fbPis.m_SetByRecipe(stPis:=stPis_OutSelect, 		req:=E_Piston_Recipe_State.Act);
fbPis.m_SetByRecipe(stPis:=stPis_OutMarinade, 		req:=E_Piston_Recipe_State.Release);
fbPis.m_SetByRecipe(stPis:=stPis_OutColor, 			req:=E_Piston_Recipe_State.Release);
fbPis.m_SetByRecipe(stPis:=stPis_Drain, 			req:=E_Piston_Recipe_State.Release);
END_ACTION

ACTION _aColor_2_entry:
fbPis.m_SetByRecipe(stPis:=stPis_Drain, 			req:=E_Piston_Recipe_State.Act);
END_ACTION

ACTION _aColor_3_active:
bStepDone:=FALSE;
IF TRUE 
AND eStatus=E_TriBlenderSelect.eColor
THEN;
	bStepDone:=TRUE;
END_IF
END_ACTION

ACTION _aColor_3_entry:
fbPis.m_SetByRecipe(stPis:=stPis_InSelect, 			req:=E_Piston_Recipe_State.Act);
fbPis.m_SetByRecipe(stPis:=stPis_InMarinade, 		req:=E_Piston_Recipe_State.Release);
fbPis.m_SetByRecipe(stPis:=stPis_InColor, 			req:=E_Piston_Recipe_State.Release);
fbPis.m_SetByRecipe(stPis:=stPis_OutSelect, 		req:=E_Piston_Recipe_State.Act);
fbPis.m_SetByRecipe(stPis:=stPis_OutMarinade, 		req:=E_Piston_Recipe_State.Release);
fbPis.m_SetByRecipe(stPis:=stPis_OutColor, 			req:=E_Piston_Recipe_State.Release);
fbPis.m_SetByRecipe(stPis:=stPis_Drain, 			req:=E_Piston_Recipe_State.Release);
END_ACTION

ACTION _aDone_entry:
eProcess:=E_TriBlenderSelect.eNone;
eReq:=E_TriBlenderSelect.eNone;
eStatus:=E_TriBlenderSelect.eNone;
bRun:=FALSE;
bDone:=TRUE;
END_ACTION

ACTION _aDrain_active:
bStepDone:=FALSE;
IF TRUE 
AND eStatus=E_TriBlenderSelect.eDrain
THEN;
	bStepDone:=TRUE;
END_IF
END_ACTION

ACTION _aDrain_entry:
fbPis.m_SetByRecipe(stPis:=stPis_InSelect, 			req:=E_Piston_Recipe_State.Release);
fbPis.m_SetByRecipe(stPis:=stPis_InMarinade, 		req:=E_Piston_Recipe_State.Act);
fbPis.m_SetByRecipe(stPis:=stPis_InColor, 			req:=E_Piston_Recipe_State.Act);
fbPis.m_SetByRecipe(stPis:=stPis_OutSelect, 		req:=E_Piston_Recipe_State.Release);
fbPis.m_SetByRecipe(stPis:=stPis_OutMarinade, 		req:=E_Piston_Recipe_State.Act);
fbPis.m_SetByRecipe(stPis:=stPis_OutColor, 			req:=E_Piston_Recipe_State.Act);
fbPis.m_SetByRecipe(stPis:=stPis_Drain, 			req:=E_Piston_Recipe_State.Act);
END_ACTION

ACTION _aInit_active:
SFCReset:=FALSE;
END_ACTION

ACTION _aMarinade_1_active:
bStepDone:=FALSE;
IF TRUE 
AND eStatus=E_TriBlenderSelect.eMarinade
THEN;
	bStepDone:=TRUE;
END_IF
END_ACTION

ACTION _aMarinade_1_entry:
fbPis.m_SetByRecipe(stPis:=stPis_InSelect, 			req:=E_Piston_Recipe_State.Release);
fbPis.m_SetByRecipe(stPis:=stPis_InMarinade, 		req:=E_Piston_Recipe_State.Release);
fbPis.m_SetByRecipe(stPis:=stPis_InColor, 			req:=E_Piston_Recipe_State.Release);
fbPis.m_SetByRecipe(stPis:=stPis_OutSelect, 		req:=E_Piston_Recipe_State.Release);
fbPis.m_SetByRecipe(stPis:=stPis_OutMarinade, 		req:=E_Piston_Recipe_State.Release);
fbPis.m_SetByRecipe(stPis:=stPis_OutColor, 			req:=E_Piston_Recipe_State.Release);
fbPis.m_SetByRecipe(stPis:=stPis_Drain, 			req:=E_Piston_Recipe_State.Release);
END_ACTION

ACTION _aMarinade_2_entry:
fbPis.m_SetByRecipe(stPis:=stPis_Drain, 			req:=E_Piston_Recipe_State.Act);
END_ACTION

ACTION _aMarinade_3_active:
bStepDone:=FALSE;
IF TRUE 
AND eStatus=E_TriBlenderSelect.eMarinade
THEN;
	bStepDone:=TRUE;
END_IF
END_ACTION

ACTION _aMarinade_3_entry:
fbPis.m_SetByRecipe(stPis:=stPis_InSelect, 			req:=E_Piston_Recipe_State.Release);
fbPis.m_SetByRecipe(stPis:=stPis_InMarinade, 		req:=E_Piston_Recipe_State.Release);
fbPis.m_SetByRecipe(stPis:=stPis_InColor, 			req:=E_Piston_Recipe_State.Release);
fbPis.m_SetByRecipe(stPis:=stPis_OutSelect, 		req:=E_Piston_Recipe_State.Release);
fbPis.m_SetByRecipe(stPis:=stPis_OutMarinade, 		req:=E_Piston_Recipe_State.Release);
fbPis.m_SetByRecipe(stPis:=stPis_OutColor, 			req:=E_Piston_Recipe_State.Release);
fbPis.m_SetByRecipe(stPis:=stPis_Drain, 			req:=E_Piston_Recipe_State.Release);
END_ACTION

ACTION _aReady_active:

eStatus:=E_TriBlenderSelect.eNone;
CASE eReq OF
	E_TriBlenderSelect.eColor:;
			IF TRUE THEN;
				eProcess:=E_TriBlenderSelect.eColor;
			END_IF	
			
	E_TriBlenderSelect.eDrain:;
			IF TRUE THEN;
				eProcess:=E_TriBlenderSelect.eDrain;
			END_IF
			
	E_TriBlenderSelect.eMarinade:;
			IF TRUE THEN;
				eProcess:=E_TriBlenderSelect.eMarinade;
			END_IF

END_CASE
END_ACTION

ACTION act_GetReference:
m_Set_SFCFlags_Reference();
//refElement REF= fbElement[eElementID];

stPis_InSelect	 REF= g_Piston.stPis[valInSelect];
stPis_InMarinade REF= g_Piston.stPis[valInMarinade];
stPis_InColor	 REF= g_Piston.stPis[valInColor];

stPis_OutSelect	  REF= g_Piston.stPis[valOutSelect];
stPis_OutMarinade REF= g_Piston.stPis[valOutMarinade];
stPis_OutColor	  REF= g_Piston.stPis[valOutColor];

stPis_Drain		  REF= g_Piston.stPis[valDrain];
END_ACTION

ACTION act_Oper:
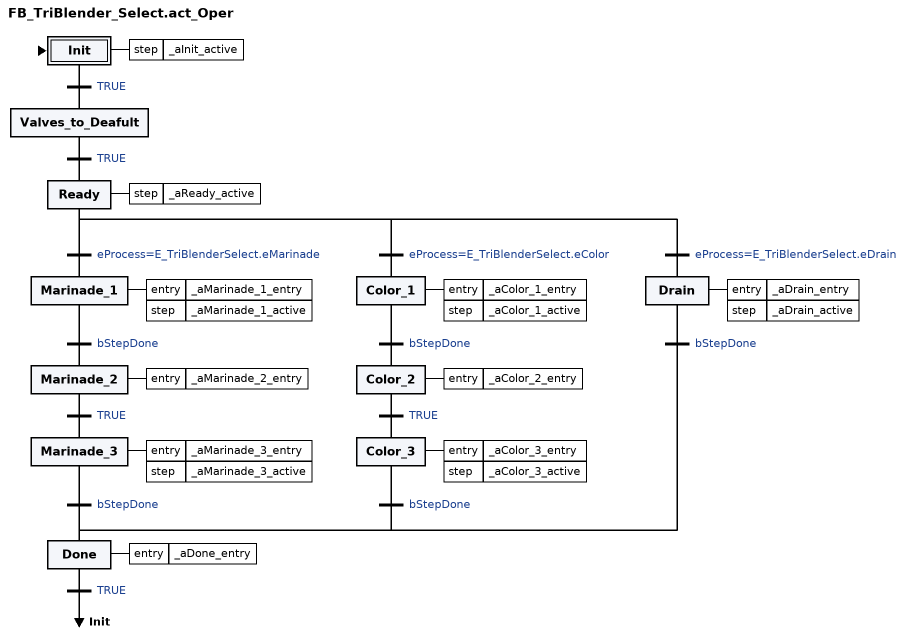
INITIAL_STEP Init:
    _aInit_active(N);  // step action
END_STEP
TRANSITION FROM Init TO Valves_to_Deafult
    := TRUE;
END_TRANSITION
STEP Valves_to_Deafult:
END_STEP
TRANSITION FROM Valves_to_Deafult TO Ready
    := TRUE;
END_TRANSITION
STEP Ready:
    _aReady_active(N);  // step action
END_STEP
TRANSITION FROM Ready TO Marinade_1
    := eProcess=E_TriBlenderSelect.eMarinade;
END_TRANSITION
STEP Marinade_1:
    _aMarinade_1_entry(P1);  // entry action
    _aMarinade_1_active(N);  // step action
END_STEP
TRANSITION FROM Marinade_1 TO Marinade_2
    := bStepDone;
END_TRANSITION
STEP Marinade_2:  // min time T#10s
    _aMarinade_2_entry(P1);  // entry action
END_STEP
TRANSITION FROM Marinade_2 TO Marinade_3
    := TRUE;
END_TRANSITION
STEP Marinade_3:
    _aMarinade_3_entry(P1);  // entry action
    _aMarinade_3_active(N);  // step action
END_STEP
TRANSITION FROM Marinade_3 TO Done
    := bStepDone;
END_TRANSITION
TRANSITION FROM Ready TO Color_1
    := eProcess=E_TriBlenderSelect.eColor;
END_TRANSITION
STEP Color_1:
    _aColor_1_entry(P1);  // entry action
    _aColor_1_active(N);  // step action
END_STEP
TRANSITION FROM Color_1 TO Color_2
    := bStepDone;
END_TRANSITION
STEP Color_2:  // min time T#10s
    _aColor_2_entry(P1);  // entry action
END_STEP
TRANSITION FROM Color_2 TO Color_3
    := TRUE;
END_TRANSITION
STEP Color_3:
    _aColor_3_entry(P1);  // entry action
    _aColor_3_active(N);  // step action
END_STEP
TRANSITION FROM Color_3 TO Done
    := bStepDone;
END_TRANSITION
TRANSITION FROM Ready TO Drain
    := eProcess=E_TriBlenderSelect.eDrain;
END_TRANSITION
STEP Drain:
    _aDrain_entry(P1);  // entry action
    _aDrain_active(N);  // step action
END_STEP
TRANSITION FROM Drain TO Done
    := bStepDone;
END_TRANSITION
STEP Done:  // min time T#0.2s
    _aDone_entry(P1);  // entry action
END_STEP
TRANSITION FROM Done TO Init
    := TRUE;
END_TRANSITION
// branch label Branch0_act_Oper_Tank
END_ACTION

ACTION act_Status:
IF TRUE 
AND fbPis.m_CheckByRecipe(stPis:=stPis_InSelect, 		req:=E_Piston_Recipe_State.Release)
AND fbPis.m_CheckByRecipe(stPis:=stPis_InMarinade, 		req:=E_Piston_Recipe_State.Release)
AND fbPis.m_CheckByRecipe(stPis:=stPis_InColor, 		req:=E_Piston_Recipe_State.Release)
AND fbPis.m_CheckByRecipe(stPis:=stPis_OutSelect, 		req:=E_Piston_Recipe_State.Release)
AND fbPis.m_CheckByRecipe(stPis:=stPis_OutMarinade, 	req:=E_Piston_Recipe_State.Release)
AND fbPis.m_CheckByRecipe(stPis:=stPis_OutColor, 		req:=E_Piston_Recipe_State.Release)
AND fbPis.m_CheckByRecipe(stPis:=stPis_Drain	, 		req:=E_Piston_Recipe_State.Release)
THEN;
	eStatus:=E_TriBlenderSelect.eMarinade;
	
ELSIF TRUE 
AND fbPis.m_CheckByRecipe(stPis:=stPis_InSelect, 		req:=E_Piston_Recipe_State.Act)
AND fbPis.m_CheckByRecipe(stPis:=stPis_InMarinade, 		req:=E_Piston_Recipe_State.Release)
AND fbPis.m_CheckByRecipe(stPis:=stPis_InColor, 		req:=E_Piston_Recipe_State.Release)
AND fbPis.m_CheckByRecipe(stPis:=stPis_OutSelect, 		req:=E_Piston_Recipe_State.Act)
AND fbPis.m_CheckByRecipe(stPis:=stPis_OutMarinade, 	req:=E_Piston_Recipe_State.Release)
AND fbPis.m_CheckByRecipe(stPis:=stPis_OutColor, 		req:=E_Piston_Recipe_State.Release)
AND fbPis.m_CheckByRecipe(stPis:=stPis_Drain	, 		req:=E_Piston_Recipe_State.Release)
THEN;
	eStatus:=E_TriBlenderSelect.eColor;
	
ELSIF TRUE 
AND fbPis.m_CheckByRecipe(stPis:=stPis_InSelect, 		req:=E_Piston_Recipe_State.Release)
AND fbPis.m_CheckByRecipe(stPis:=stPis_InMarinade, 		req:=E_Piston_Recipe_State.Act)
AND fbPis.m_CheckByRecipe(stPis:=stPis_InColor, 		req:=E_Piston_Recipe_State.Act)
AND fbPis.m_CheckByRecipe(stPis:=stPis_OutSelect, 		req:=E_Piston_Recipe_State.Release)
AND fbPis.m_CheckByRecipe(stPis:=stPis_OutMarinade, 	req:=E_Piston_Recipe_State.Act)
AND fbPis.m_CheckByRecipe(stPis:=stPis_OutColor, 		req:=E_Piston_Recipe_State.Act)
AND fbPis.m_CheckByRecipe(stPis:=stPis_Drain	, 		req:=E_Piston_Recipe_State.Act)
THEN;
	eStatus:=E_TriBlenderSelect.eDrain;
	
ELSE
	eStatus:=E_TriBlenderSelect.eNone;
	
END_IF;
END_ACTION

METHOD m_CheckStatus : BOOL
VAR_INPUT
	eReqStatus		: E_TriBlenderSelect;
END_VAR
IF eStatus=eReqStatus 
AND eProcess=E_TriBlenderSelect.eNone
AND eReq=E_TriBlenderSelect.eNone
AND bReady
AND bDone
AND NOT bRun
THEN;
	m_CheckStatus:=TRUE;
END_IF
END_METHOD

METHOD m_Request_Reset : BOOL
VAR_IN_OUT
	memo: R_TRIG;
END_VAR
memo(CLK:=eReq=0);
IF TRUE 
AND memo.Q
THEN;
	SFCReset:=TRUE;
END_IF
END_METHOD

METHOD m_Run : BOOL
VAR_INPUT
	eReqProc			: E_TriBlenderSelect;
END_VAR
IF eProcess=E_TriBlenderSelect.eNone THEN;
	eProcess:=eReq:=eReqProc;
	bDone:=FALSE;
	m_Run:=TRUE;
END_IF
END_METHOD

METHOD m_Set_Request : BOOL
VAR_INPUT
	eSetReg		: E_TriBlenderSelect;
END_VAR
eReq:=eSetReg;
END_METHOD

{warning 'add method implementation '}
METHOD m_Set_SFCFlags_Reference : BOOL
//Set reference to SFC flags

refSFC.SFCInit REF= SFCInit;
refSFC.SFCReset REF= SFCReset;
refSFC.SFCError REF= SFCError;
refSFC.SFCEnableLimit REF= SFCEnableLimit;
refSFC.SFCErrorStep REF= SFCErrorStep;
refSFC.SFCErrorPOU REF= SFCErrorPOU;
refSFC.SFCQuitError REF= SFCQuitError;
refSFC.SFCPause REF= SFCPause;
refSFC.SFCTrans REF= SFCTrans;
refSFC.SFCCurrentStep REF= SFCCurrentStep;
refSFC.SFCTip REF= SFCTip;
refSFC.SFCTipMode REF= SFCTipMode;

// Cycle handle for SFC
m_SFC_Handle();
END_METHOD

END_FUNCTION_BLOCK

// ---- 03 Project/12 TriBlender/FB_Dissolving.TcPOU
FUNCTION_BLOCK PUBLIC FB_Dissolving EXTENDS FB_SFC_Cycle IMPLEMENTS ITF_FB_SFC_Cycle
VAR_INPUT
END_VAR
VAR_OUTPUT
END_VAR
VAR
	step: INT;
	i: INT;
	ton_Blending_Speed: TON;
	tBlending: TIME;
	tBlending_count: TIME;
	ptTemp: DINT;
	tBlendingRemainTime: DINT;
	realTemp: REAL;
	fBlendingPercenatge: DINT;
END_VAR

VAR_IN_OUT
	fb_TriBlender			: FB_Pump;
END_VAR

m_Set_SFCFlags_Reference();
act_Oper();
IF g_HMI_Panel.stPLC_To_VisuPLC.iActual_Component<>0 THEN
	ptTemp:=TIME_TO_DINT(g_HMI_Panel.stPLC_To_VisuPLC.arr_Component[g_HMI_Panel.stPLC_To_VisuPLC.iActual_Component].tBlendingDuration);
ELSE;
	ptTemp:=0;
END_IF

tBlendingRemainTime:=ptTemp - TIME_TO_DINT(tBlending);
IF ptTemp<>0 THEN;
	realTemp:=(DINT_TO_REAL(tBlendingRemainTime)/DINT_TO_REAL(ptTemp)*100.0);
	fBlendingPercenatge:=TRUNC(realTemp);
END_IF

ACTION _aChek_if_Done_active:
bStepDone:=FALSE;
IF g_HMI_Panel.stPLC_To_VisuPLC.iActual_Component >= 10 THEN;
	bStepDone:=TRUE;
END_IF
END_ACTION

ACTION _aComponent_Blending_active:
bStepDone:=FALSE;
IF tBlending > g_HMI_Panel.stPLC_To_VisuPLC.arr_Component[g_HMI_Panel.stPLC_To_VisuPLC.iActual_Component].tBlendingDuration THEN;
	bStepDone:=TRUE;
	g_HMI_Panel.stPLC_To_VisuPLC.bBlending_Active:=FALSE;
END_IF

fb_TriBlender.m_Run(RPM:=g_HMI_Panel.stPLC_To_VisuPLC.arr_Component[g_HMI_Panel.stPLC_To_VisuPLC.iActual_Component].rFlowRate_Blending);

ton_Blending_Speed(PT:=T#2S);
IF TRUE 
AND fb_TriBlender.m_Get_Speed() >= g_HMI_Panel.stPLC_To_VisuPLC.arr_Component[g_HMI_Panel.stPLC_To_VisuPLC.iActual_Component].rFlowRate_Blending - 10
AND fb_TriBlender.m_Get_Speed() <= g_HMI_Panel.stPLC_To_VisuPLC.arr_Component[g_HMI_Panel.stPLC_To_VisuPLC.iActual_Component].rFlowRate_Blending + 10
THEN;
	ton_Blending_Speed.IN:=TRUE;
ELSE;
	ton_Blending_Speed.IN:=FALSE;
END_IF

IF ton_Blending_Speed.Q THEN;
	tBlending:=tBlending + T#10MS; // scan Time
ELSE;
	
END_IF
END_ACTION

ACTION _aComponent_Blending_entry:
g_HMI_Panel.stPLC_To_VisuPLC.bDissolving_Active:=FALSE;
g_HMI_Panel.stPLC_To_VisuPLC.bBlending_Active:=TRUE;
END_ACTION

ACTION _aDissolving_Done_entry:
bDisolvingProcess_Done:=TRUE;
END_ACTION

ACTION _aInit_Dissolve_exit:
step:=0;
g_HMI_Panel.stPLC_To_VisuPLC.iActual_Component:=0;
g_HMI_Panel.stPLC_To_VisuPLC.bDissolving_Active:=FALSE;
g_HMI_Panel.stPLC_To_VisuPLC.bBlending_Active:=FALSE;
bRun:=FALSE;
END_ACTION

ACTION _aReady_exit:
g_HMI_Panel.stPLC_To_VisuPLC.iActual_Component:=1;
g_HMI_Panel.stPLC_To_VisuPLC.bDissolving_Active:=FALSE;
END_ACTION

ACTION _arepeat_stage_active:
bStepDone:=NOT g_HMI_Panel.stVisuPLC_To_PLC.bActualComponentDisolving_Done;
END_ACTION

ACTION _aSet_Next_Component_active:
bStepDone:=FALSE;
IF g_HMI_Panel.stVisuPLC_To_PLC.bActualComponentDisolving_Done THEN;
	bStepDone:=TRUE;
END_IF

IF g_HMI_Panel.stVisuPLC_To_PLC.bPauseTriBlender THEN;
	fb_TriBlender.m_Stop();
ELSE;
	fb_TriBlender.m_Run(RPM:=g_HMI_Panel.stVisuPLC_To_PLC.RPM_setPoint);
END_IF
END_ACTION

ACTION _aSet_Next_Component_entry:
g_HMI_Panel.stPLC_To_VisuPLC.bDissolving_Active:=FALSE;
g_HMI_Panel.stPLC_To_VisuPLC.bBlending_Active:=FALSE;
g_HMI_Panel.stPLC_To_VisuPLC.iActual_Component:=g_HMI_Panel.stPLC_To_VisuPLC.iActual_Component+1;

FOR i:=g_HMI_Panel.stPLC_To_VisuPLC.iActual_Component TO 10 DO
	IF g_HMI_Panel.stPLC_To_VisuPLC.arr_Component[i].rWeight>0 THEN;
		g_HMI_Panel.stPLC_To_VisuPLC.iActual_Component:=i;
		g_HMI_Panel.stPLC_To_VisuPLC.bDissolving_Active:=TRUE;
		EXIT;
	END_IF
END_FOR

tBlending:=T#0S;
END_ACTION

ACTION act_Oper:
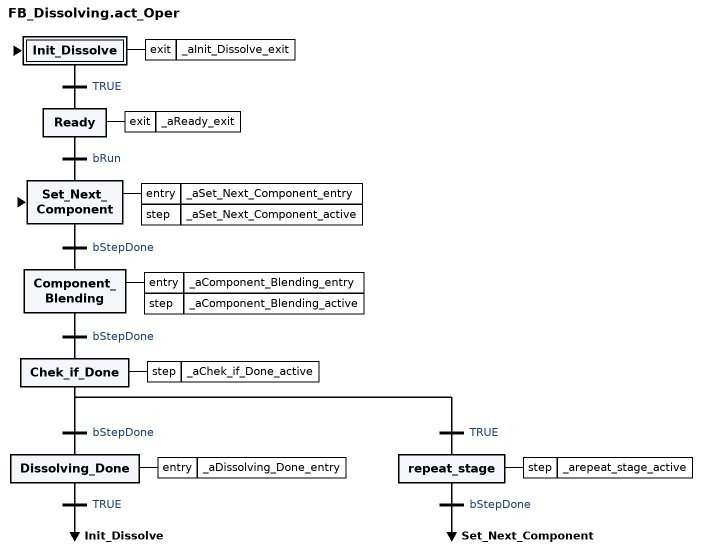
INITIAL_STEP Init_Dissolve:
    _aInit_Dissolve_exit(P0);  // exit action
END_STEP
TRANSITION FROM Init_Dissolve TO Ready
    := TRUE;
END_TRANSITION
STEP Ready:
    _aReady_exit(P0);  // exit action
END_STEP
TRANSITION FROM Ready TO Set_Next_Component
    := bRun;
END_TRANSITION
STEP Set_Next_Component:
    _aSet_Next_Component_entry(P1);  // entry action
    _aSet_Next_Component_active(N);  // step action
END_STEP
TRANSITION FROM Set_Next_Component TO Component_Blending
    := bStepDone;
END_TRANSITION
STEP Component_Blending:
    _aComponent_Blending_entry(P1);  // entry action
    _aComponent_Blending_active(N);  // step action
END_STEP
TRANSITION FROM Component_Blending TO Chek_if_Done
    := bStepDone;
END_TRANSITION
STEP Chek_if_Done:
    _aChek_if_Done_active(N);  // step action
END_STEP
TRANSITION FROM Chek_if_Done TO Dissolving_Done
    := bStepDone;
END_TRANSITION
TRANSITION FROM Chek_if_Done TO repeat_stage
    := TRUE;
END_TRANSITION
STEP repeat_stage:
    _arepeat_stage_active(N);  // step action
END_STEP
TRANSITION FROM repeat_stage TO Set_Next_Component
    := bStepDone;
END_TRANSITION
STEP Dissolving_Done:
    _aDissolving_Done_entry(P1);  // entry action
END_STEP
TRANSITION FROM Dissolving_Done TO Init_Dissolve
    := TRUE;
END_TRANSITION
// branch label Branch0_act_Oper
END_ACTION

METHOD m_Set_SFCFlags_Reference : BOOL
//Set reference to SFC flags

refSFC.SFCInit REF= SFCInit;
refSFC.SFCReset REF= SFCReset;
refSFC.SFCError REF= SFCError;
refSFC.SFCEnableLimit REF= SFCEnableLimit;
refSFC.SFCErrorStep REF= SFCErrorStep;
refSFC.SFCErrorPOU REF= SFCErrorPOU;
refSFC.SFCQuitError REF= SFCQuitError;
refSFC.SFCPause REF= SFCPause;
refSFC.SFCTrans REF= SFCTrans;
refSFC.SFCCurrentStep REF= SFCCurrentStep;
refSFC.SFCTip REF= SFCTip;
refSFC.SFCTipMode REF= SFCTipMode;

// Cycle handle for SFC
m_SFC_Handle();
END_METHOD

END_FUNCTION_BLOCK

// ---- 03 Project/13 Weight control/WeighingModule/Rs232Logging.TcPOU
PROGRAM Rs232Logging
VAR


	fbPcCom		: FB_SerialCom;
	
	(* exchange buffers with background communication with the PC COM port device *)
	RxBufferPcCom	: ComBuffer;	(* Receive data buffer; used with all receive function blocks *)
	TxBufferPcCom	: ComBuffer;	(* Transmit data buffer; used with all receive function blocks *)
	
END_VAR

VAR_OUTPUT
	rWeight: REAL;
END_VAR




(* background communication with the PC COM port device *)
BackgroundPcCOM(RxBufferPcCom:=RxBufferPcCom, TxBufferPcCom:=TxBufferPcCom);


(* Send and receive commands *)
fbPcCom(TxBuffer:=TxBufferPcCom, RxBuffer:=RxBufferPcCom);
	
 rWeight:=fbPcCom.Weight;

END_PROGRAM

// ---- 03 Project/13 Weight control/WeighingModule/FB_SerialCom.TcPOU
FUNCTION_BLOCK FB_SerialCom
VAR_IN_OUT
	TxBuffer	: ComBuffer;
	RxBuffer	: ComBuffer;
END_VAR
VAR
	Timer		: TON := (PT:=T#1S);
	fbSend		: SendString;
	bSendBusy	: BOOL;
	eSendErrorID: ComError_t;

	fbReceive		: ReceiveString;
	sReceivedString	: STRING;
	sLastReceivedString: STRING;
	bStringReceived	: BOOL;
	bReceiveBusy	: BOOL;
	bReceiveError	: BOOL;
	eReceiveErrorID	: ComError_t;
	bReceiveTimeout	: BOOL;
	nReceiveCounter	: UDINT;
	
	Prefix: STRING;
	Suffix: STRING;
	NotReceive: INT;
END_VAR
VAR_OUTPUT
	Weight: REAL;
END_VAR

// Call the send block every second to repeat the transmission.
// Also call the block as long as it is busy to finish a transmission.
(*Timer(IN:=TRUE);
IF Timer.Q OR fbSend.Busy THEN
	Timer(IN:=FALSE); (* reset timer *)
	fbSend(	SendString:= '$02Hello World ! $03',
			TXbuffer:= TxBuffer,
			Busy=> bSendBusy,
			Error=> );
	IF fbSend.Error <> COMERROR_NOERROR THEN
		eSendErrorID := fbSend.Error;
	END_IF
END_IF*)

//	Receive string data:
//	The block receives any data strings beginning with a STX ($02) and ending with an ETX ($03) character.	
fbReceive(
	Prefix:= Prefix,//'$02',
	Suffix:=Suffix,//'$R$N', //'$03'
	Timeout:= T#1s,
	ReceivedString:= sReceivedString,
	RXbuffer:= RxBuffer,
	StringReceived=> bStringReceived,
	Busy=> bReceiveBusy,
	Error=> ,
	RxTimeout=> bReceiveTimeout );
IF fbReceive.Error <> COMERROR_NOERROR THEN
	eReceiveErrorID := fbReceive.Error;
END_IF
IF bStringReceived THEN
	nReceiveCounter := nReceiveCounter + 1;
	sLastReceivedString := sReceivedString;
ELSE
	NotReceive:= NotReceive+1;
	
END_IF

Weight:= STRING_TO_REAL(sLastReceivedString);

END_FUNCTION_BLOCK

// ---- 03 Project/13 Weight control/WeighingModule/BackgroundPcCOM.TcPOU
PROGRAM BackgroundPcCOM
VAR_IN_OUT
	RxBufferPcCom		: ComBuffer;	(* Receive data buffer; used with all receive function blocks *)
	TxBufferPcCom		: ComBuffer;	(* Transmit data buffer; used with all receive function blocks *)
END_VAR
VAR
	(* background communication with the PC COM port device *)
	fbPcComCtrl			: SerialLineControl;
	bPcComCtrlError		: BOOL;
	ePcComCtrlErrorID	: ComError_t;	
	(* 	I/O variables for a PC-COM port *)
	stIn_PcCom AT %I*	: EL6inData22B;	(* linked to the port in the TwinCAT System Manager *)
	stOut_PcCom AT %Q*	: EL6outData22B;	(* linked to the port in the TwinCAT System Manager *)
	ComMode: ComSerialLineMode_t := COMSERIALLINEMODE_T.SERIALLINEMODE_EL6_22B;
END_VAR

(*
The SerialLineControl function block is supposed to be called in every PLC cycle.
It communicates with the serial line hardware device and transmits or receives data.
The SerialLineControl can be called in the standard task (e.g.for PcCOM port usage) 
or in a separate fast task (e.g.for terminal usage) as well.
A fast separate task will be necessary at high baud rates or with KL6001 terminals 
which have a small process image (3 or 5 data bytes only)
*)

(* background communication with the PC COM port device *)
fbPcComCtrl(
	Mode:= ComMode,//SERIALLINEMODE_PC_COM_PORT, 
	pComIn:= ADR(stIn_PcCom), 
	pComOut:= ADR(stOut_PcCom), 
	SizeComIn:= SIZEOF(stIn_PcCom), 
	Error=> , 
	ErrorID=> , 
	TxBuffer:= TxBufferPcCom, 
	RxBuffer:= RxBufferPcCom );
IF fbPcComCtrl.Error THEN
	bPcComCtrlError := TRUE;
	ePcComCtrlErrorID := fbPcComCtrl.ErrorID;
END_IF

END_PROGRAM

// ---- 03 Project/12 TriBlender/prg_PLCs_communication.TcPOU
PROGRAM prg_PLCs_communication
VAR
	fbAdsRead: ADSREAD;
	fbAdsWrite: ADSWRITE;

	ton_Update: TON;
END_VAR

ton_Update(PT:=T#50MS, IN:=NOT ton_Update.Q);

IF ton_Update.Q THEN;
END_IF	

fbAdsRead(
	NETID:= , 
	PORT:= 852, 
	IDXGRP:= 16#4020,// 
	IDXOFFS:= 1000,// 
	LEN:= SIZEOF(g_HMI_Panel.stVisuPLC_To_PLC), 
	DESTADDR:= ADR(g_HMI_Panel.stVisuPLC_To_PLC), 
	READ:= ton_Update.Q, 
	TMOUT:= , 
	BUSY=> , 
	ERR=> , 
	ERRID=> );
	
fbAdsWrite(
	NETID:= , 
	PORT:= 852, 
	IDXGRP:= 16#4020,// 
	IDXOFFS:= 2000, //
	LEN:= SIZEOF(g_HMI_Panel.stPLC_To_VisuPLC), 
	SRCADDR:= ADR(g_HMI_Panel.stPLC_To_VisuPLC), 
	WRITE:= ton_Update.Q, 
	TMOUT:= , 
	BUSY=> , 
	ERR=> , 
	ERRID=> );
	
g_HMI_Panel.stPLC_To_VisuPLC.lifeBit:=NOT g_HMI_Panel.stVisuPLC_To_PLC.lifeBit;

act_Send_To_HMI();
act_Get_From_HMI();

ACTION act_Get_From_HMI:

END_ACTION

ACTION act_Send_To_HMI:


CASE eTriBlenderUsage OF
	E_TriBlenderUsage.eMarinada_T1:;
		(*g_HMI_Panel.q_stPLC_To_VisuPLC.Description:=fbTank1.stProdParam.stRecipe.Description;
		g_HMI_Panel.q_stPLC_To_VisuPLC.prodType:=fbTank1.stProdParam.stRecipe.prodType;
		g_HMI_Panel.q_stPLC_To_VisuPLC.arr_Component:=fbTank1.stProdParam.stRecipe.arr_Component;
		g_HMI_Panel.q_stPLC_To_VisuPLC.:=fbTank1.stProdParam.stRecipe.Description;*)
		m_GetProductionInfo(fbProductionTank:=fbTank1);		
	E_TriBlenderUsage.eMarinada_T2:;
		m_GetProductionInfo(fbProductionTank:=fbTank2);
	E_TriBlenderUsage.eColor_T3:;
		m_GetProductionInfo(fbProductionTank:=fbTank3);
	E_TriBlenderUsage.eColor_T4:;
		m_GetProductionInfo(fbProductionTank:=fbTank4);
		
ELSE;
	
	m_CleanProductionInfo();
END_CASE

g_HMI_Panel.stPLC_To_VisuPLC.RPM_FeedBack:=g_Pump.fbPump[E_Pump_List.TB0001].m_Get_Speed();
g_HMI_Panel.stPLC_To_VisuPLC.Flow_FeedBack:=g_AnalogSensor.stAnalogSensor[E_ASense_Name.FT9012].Value;
g_HMI_Panel.stPLC_To_VisuPLC.fBlendingPercenatge:=fbDissolving.fBlendingPercenatge;

CASE g_Data.eTriBlenderUsage OF
	E_TriBlenderUsage.eMarinada_T1,E_TriBlenderUsage.eMarinada_T2:;
			g_HMI_Panel.stPLC_To_VisuPLC.bMainPause_Active:=stOper[E_ModeZone.eTriBlender_Marinade].iActOperation=E_OperationButtons.ePauseAll;
	E_TriBlenderUsage.eColor_T3,E_TriBlenderUsage.eColor_T4:;
			g_HMI_Panel.stPLC_To_VisuPLC.bMainPause_Active:=stOper[E_ModeZone.eTriBlender_Color].iActOperation=E_OperationButtons.ePauseAll;
END_CASE
END_ACTION

METHOD m_CleanProductionInfo : BOOL
VAR
	stRecipe_Clean: ST_Prod_Recipe;	
	i: INT;
END_VAR

g_HMI_Panel.stPLC_To_VisuPLC.Description:='Not Loaded';
//g_HMI_Panel.stPLC_To_VisuPLC.prodType:=E_Prod_Type.Marinade;
FOR i:=1 TO 10 DO
	stRecipe_Clean.arr_Component[i].sDescription:='-*-*-';
END_FOR
g_HMI_Panel.stPLC_To_VisuPLC.arr_Component:=stRecipe_Clean.arr_Component;
END_METHOD

METHOD m_GetProductionInfo : BOOL
VAR_INPUT
	fbProductionTank: FB_ProductionTank;
END_VAR
g_HMI_Panel.q_stPLC_To_VisuPLC.Description:=fbProductionTank.stProdParam.stRecipe.Description;
g_HMI_Panel.q_stPLC_To_VisuPLC.prodType:=fbProductionTank.stProdParam.stRecipe.prodType;
g_HMI_Panel.q_stPLC_To_VisuPLC.arr_Component:=fbProductionTank.stProdParam.stRecipe.arr_Component;
		
g_HMI_Panel.stPLC_To_VisuPLC.Description:=fbProductionTank.stProdParam.stRecipe.Description;
g_HMI_Panel.stPLC_To_VisuPLC.prodType:=fbProductionTank.stProdParam.stRecipe.prodType;
g_HMI_Panel.stPLC_To_VisuPLC.arr_Component:=fbProductionTank.stProdParam.stRecipe.arr_Component;
END_METHOD

END_PROGRAM

// ---- 00 Library/04 Recipe/FB_Recipe.TcPOU
FUNCTION_BLOCK FB_Recipe
VAR_INPUT
	pstRecipe				:POINTER TO ST_Recipe;
	bMemoRecipeUpdated		:BOOL:=FALSE;
	sRecipeDef				:STRING; (* current recipe definition *)
	bLoadDefault			:BOOL;
	sRecipesStoragePath		:STRING;
	bHMI_FrameActive		:BOOL;

END_VAR

VAR
	i						:INT;	
	RecipeManCommands 		:RecipeManCommands; (* Recipe Manager *)
	k						:INT;
	t1						:TON;
	check					:DWORD;
	INDEX					:INT:= 0;
	bReloadRecipes			:BOOL;
	rt_LoadDefault: R_TRIG;
	MessageBox			:MessageBox_Struct;
	arrLastReturn		: ARRAY[0..15] OF DWORD;
	LastReturn			:  DWORD;
	ton_RecipeUpdated: TON;
	sMessage: STRING;
	ton_SetStoragePath_Delay: TON;
	bSetStoragePath: BOOL:=TRUE;
	ton_SetStoragePathTimeOut: TON;
	bReturn: BOOL;
	
	ton_MessClear: TON;
	rt_Init: R_TRIG;
	sLastMessage: STRING;
	rt_Saved: R_TRIG;
	rt_FrameAvtive: R_TRIG;
	rt_LoadDefault1: R_TRIG;
END_VAR

act_SetStoragePath();
act_Disp();

IF pstRecipe^.bValidSelected THEN
	pstRecipe^.sSelectedReceipe:= pstRecipe^.arrRecipeNames[pstRecipe^.iRecipeIndex];
	pstRecipe^.bValidSelected:=FALSE;
END_IF

rt_FrameAvtive(CLK:=bHMI_FrameActive);
rt_LoadDefault1(CLK:=bLoadDefault);
IF pstRecipe^.bReInit OR rt_LoadDefault1.Q OR rt_FrameAvtive.Q THEN;
	pstRecipe^.bReInit:=FALSE;
	pstRecipe^.bInit:=FALSE;
	bSetStoragePath:=TRUE;
END_IF

t1(IN:=NOT pstRecipe^.bInit , PT:=T#0.5S);
IF (NOT pstRecipe^.bInit AND t1.Q) THEN
	
	IF NOT bSetStoragePath THEN;
		arrLastReturn[3]:=RecipeManCommands.ResetLastInfo();
		arrLastReturn[4]:=RecipeManCommands.ReloadRecipes(RecipeDefinitionName:=sRecipeDef);
		pstRecipe^.iRecipeCount:=RecipeManCommands.GetRecipeCount(sRecipeDef);
		FOR i := 0 TO GVL_Recipe.C_Max_RecipeFileNum DO
			pstRecipe^.arrRecipeNames[i] := '';
		END_FOR
		FOR i := 0 TO 1200 DO
			pstRecipe^.arrVariableNamesValue[i] := '';
			pstRecipe^.arrVariableValue[i] := '';
		END_FOR	
		(* save all recipe names of one recipe definition in an array *)
		arrLastReturn[0]:=RecipeManCommands.GetRecipeNames(sRecipeDef, ADR(pstRecipe^.arrRecipeNames),GVL_Recipe.C_Max_RecipeFileNum, 0);
		pstRecipe^.iRecipeIndex:=0;
		pstRecipe^.sLastSelectedReceipe:=pstRecipe^.sSelectedReceipe:=pstRecipe^.arrRecipeNames[0];
		pstRecipe^.bInit:=TRUE;
		pstRecipe^.bReInit:=FALSE;		
	END_IF

END_IF


rt_Init(CLK:=pstRecipe^.bInit);
IF pstRecipe^.bInit THEN

	IF pstRecipe^.sSelectedReceipe <> pstRecipe^.sLastSelectedReceipe 
	OR rt_Init.Q 
	OR rt_Saved.Q
	THEN;
				 
		arrLastReturn[1]:=RecipeManCommands.GetRecipeValues
			(
			RecipeDefinitionName:= sRecipeDef,
			RecipeName:= pstRecipe^.sSelectedReceipe, 
			pStrings:= ADR(pstRecipe^.arrVariableValue), 
			iSize:= 1200, 
			iStartIndex:= 0, 
			iStringLength:=80
			 );		
					
		arrLastReturn[2]:=RecipeManCommands.GetRecipeVariableNames
			(
			RecipeDefinitionName:=sRecipeDef,
			RecipeName:=pstRecipe^.sSelectedReceipe, 
			pStrings:= ADR(pstRecipe^.arrVariableNamesValue), 
			iSize:= 1200, 
			iStartIndex:= 0
			);
				
			pstRecipe^.bShowFile:=FALSE;
	END_IF
	pstRecipe^.sLastSelectedReceipe:=pstRecipe^.sSelectedReceipe;
END_IF


FOR i:=0 TO 15 DO
	IF arrLastReturn[i]<>0 THEN
		LastReturn:=arrLastReturn[i];
		EXIT;
	END_IF
	IF i=15 AND arrLastReturn[i]=0 THEN
		LastReturn:=0;
	END_IF
END_FOR

act_Cmd_List();

ACTION act_Cmd_List:
rt_LoadDefault(CLK:=bLoadDefault AND NOT bSetStoragePath);
IF rt_LoadDefault.Q THEN;
	pstRecipe^.sSelectedReceipe:='Default';
	pstRecipe^.bWriteToPLC_Cmd:=TRUE;
END_IF


IF pstRecipe^.bReloadRecipes THEN
	arrLastReturn[3]:=RecipeManCommands.ResetLastInfo();
	arrLastReturn[4]:=RecipeManCommands.ReloadRecipes(RecipeDefinitionName:=sRecipeDef);
	pstRecipe^.bReloadRecipes:=FALSE;
END_IF


IF pstRecipe^.bGetLastError THEN
	arrLastReturn[5]:=RecipeManCommands.GetLastError();
	pstRecipe^.bGetLastError:=FALSE;
END_IF


IF pstRecipe^.bResetLastError THEN
	arrLastReturn[6]:=RecipeManCommands.ResetLastError();
	pstRecipe^.bResetLastError:=FALSE;
	sMessage:='';
	FOR i:=0 TO 15 DO
		arrLastReturn[i]:=0;
	END_FOR	
END_IF

rt_Saved(CLK:=NOT pstRecipe^.bSaveFileCmd);
IF pstRecipe^.bSaveFileCmd  THEN
	sMessage:='cmd Save Recipe';
	IF  METH_Search(pstRecipe:=pstRecipe , sSearchRecipe:=pstRecipe^.sSelectedReceipe ) THEN
		//arrLastReturn[7]:=RecipeManCommands.ReadAndSaveRecipeAs(RecipeDefinitionName:=sRecipeDef,
		arrLastReturn[7]:=RecipeManCommands.ReadAndSaveRecipe(RecipeDefinitionName:=sRecipeDef,
			RecipeName:=pstRecipe^.sSelectedReceipe);// ,
			//FileName:='.txtrecipe' );
		sMessage:='cmd Save Recipe - Done';
		pstRecipe^.bSaveFileCmd:=FALSE;
	ELSE;
		sMessage:='cmd Save Recipe - Failed';
	END_IF
END_IF


IF pstRecipe^.bWriteToPLC_Cmd  THEN
	sMessage:='cmd Load Recipe';
	bMemoRecipeUpdated:=FALSE;
	IF  METH_Search(pstRecipe:=pstRecipe , sSearchRecipe:=pstRecipe^.sSelectedReceipe ) THEN
		arrLastReturn[8]:=RecipeManCommands.LoadRecipe(RecipeDefinitionName:= sRecipeDef, RecipeName:= pstRecipe^.sSelectedReceipe);
		arrLastReturn[9]:=RecipeManCommands.WriteRecipe(RecipeDefinitionName:= sRecipeDef, RecipeName:= pstRecipe^.sSelectedReceipe);
		sMessage:='cmd Load Recipe - Done';
		pstRecipe^.bWriteToPLC_Cmd:=FALSE;
		ton_RecipeUpdated.IN:=TRUE;
	ELSE;
		sMessage:='cmd Load Recipe - Failed';
	END_IF
END_IF
ton_RecipeUpdated(PT:=T#1S);
IF ton_RecipeUpdated.Q THEN;
	bMemoRecipeUpdated:=TRUE;	
	ton_RecipeUpdated.IN:=FALSE;
END_IF


IF pstRecipe^.bCreateRecipe AND pstRecipe^.sNewRecipeName <> '' THEN
	arrLastReturn[10]:=RecipeManCommands.CreateRecipe(sRecipeDef ,pstRecipe^.sNewRecipeName);
	sMessage:='cmd Create Recipe - Done';
	pstRecipe^.bCreateRecipe:=FALSE;
	pstRecipe^.bReInit:=TRUE;
END_IF


IF pstRecipe^.bDeleteRecipe THEN
	sMessage:='cmd Delete Recipe';
	IF  METH_Search(pstRecipe:=pstRecipe , sSearchRecipe:=pstRecipe^.sSelectedReceipe ) THEN
		arrLastReturn[11]:=RecipeManCommands.DeleteRecipe(sRecipeDef ,pstRecipe^.sSelectedReceipe);
		sMessage:='cmd Delete Recipe - Done';
		pstRecipe^.bDeleteRecipe:=FALSE;
		pstRecipe^.bReInit:=TRUE;
	ELSE;
		sMessage:='cmd Delete Recipe - Failed';
	END_IF
END_IF

ton_MessClear(PT:=T#30S);
IF sMessage<>sLastMessage THEN;
	ton_MessClear(IN:=FALSE);
	sLastMessage:=sMessage;
ELSIF sMessage<>'' THEN;
	ton_MessClear.IN:=TRUE;
ELSE;
	ton_MessClear.IN:=FALSE;
END_IF
IF ton_MessClear.Q THEN;
	sMessage:='';
END_IF
END_ACTION

ACTION act_Disp:

IF pstRecipe^.iDispSel<0 THEN; pstRecipe^.iDispSel:=0; END_IF
IF pstRecipe^.iDispSel>1180 THEN; pstRecipe^.iDispSel:=1180; END_IF

//FOR k:=iDispSel TO iDispSel+19 DO;
FOR k:=0 TO 20 DO;
	pstRecipe^.arrVariableDisp[0,k]:= INT_TO_STRING(pstRecipe^.iDispSel+k);
	pstRecipe^.arrVariableDisp[1,k]:=pstRecipe^.arrVariableNamesValue[pstRecipe^.iDispSel+k];
	pstRecipe^.arrVariableDisp[2,k]:=pstRecipe^.arrVariableValue[pstRecipe^.iDispSel+k];
END_FOR
END_ACTION

ACTION act_SetStoragePath:
ton_SetStoragePath_Delay(PT:=T#0.5S,IN:=bSetStoragePath);
ton_SetStoragePathTimeOut(PT:=T#2S);

IF ton_SetStoragePath_Delay.Q THEN;
	bReturn:=RecipeManCommands.SetStoragePath(stPath:=sRecipesStoragePath);
	//sMessage:='cmd Set Storage Path';
	IF bReturn THEN;
		bSetStoragePath:=FALSE;
		ton_SetStoragePathTimeOut.IN:=FALSE;
		//sMessage:='cmd Set Storage Path - Done';
	ELSE
		ton_SetStoragePathTimeOut.IN:=TRUE;
	END_IF
	
	IF ton_SetStoragePathTimeOut.Q THEN;
		bSetStoragePath:=FALSE;
		ton_SetStoragePathTimeOut.IN:=FALSE;
		//sMessage:='cmd Set Storage Path - Failed';		
	END_IF
END_IF
END_ACTION

METHOD METH_Search : BOOL
VAR_INPUT
	pstRecipe :POINTER TO ST_Recipe;
	sSearchRecipe	:STRING(30);
END_VAR

VAR
	i: INT;
END_VAR
METH_Search:=FALSE;
FOR i:= 0 TO GVL_Recipe.C_Max_RecipeFileNum DO
	IF sSearchRecipe = pstRecipe^.arrRecipeNames[i] THEN
		METH_Search:=TRUE;
		EXIT;
	END_IF
END_FOR
END_METHOD

END_FUNCTION_BLOCK

// ---- 00 Library/04-Messages/FB_PrintErrMessageByID.TcPOU
FUNCTION_BLOCK FB_PrintErrMessageByID
VAR_INPUT
	sActErrorID			: STRING;
	iFB_Num				: INT:=0;
	sModuleDescription	:STRING:='';
END_VAR
VAR_OUTPUT
END_VAR
VAR
	cFound				: INT;
	i					: INT;
	iFound				: INT;
	bNewMeasege			: BOOL;
	rtrig1				: R_TRIG;
	sLastErrorID		: STRING;
	j: INT;
	sFB_Num: STRING(3);

END_VAR




	
	IF sActErrorID<>'000x000x000'  AND sActErrorID<>'' THEN
		IF iFB_Num>0 THEN;
			sFB_Num:=F_iFB_Num_sFB_Num(iFB_Num:=iFB_Num);
			sLastErrorID:=REPLACE(sActErrorID,sFB_Num,3,5);
		ELSE;
			sLastErrorID:=sActErrorID;
		END_IF			
		
		bNewMeasege:=TRUE;
		FOR i:=1 TO 100 DO
			IF Buffer_Act_Message[i].sErrID=sLastErrorID THEN;//sActErrorID
				//IF Buffer_Act_Message[i].sModuleDescription = sFB_ModuleDescription THEN
					bNewMeasege:=FALSE;
					EXIT; 
				//END_IF
			END_IF
		END_FOR
	ELSE
		bNewMeasege:=FALSE;
	END_IF
	
	IF bNewMeasege THEN;
		FOR i:=100 TO 2 BY -1 DO
			Buffer_Act_Message[i].sDateTime:=Buffer_Act_Message[i-1].sDateTime;
			Buffer_Act_Message[i].sErrID:=Buffer_Act_Message[i-1].sErrID;
			Buffer_Act_Message[i].sErrorMessage:=Buffer_Act_Message[i-1].sErrorMessage;
			Buffer_Act_Message[i].sLevel:=Buffer_Act_Message[i-1].sLevel;
			Buffer_Act_Message[i].sModuleDescription:=Buffer_Act_Message[i-1].sModuleDescription;
		END_FOR
		
		Buffer_Act_Message[1].sDateTime:=prg_RealClock.sRealTime_Date;
		Buffer_Act_Message[1].sErrID:=sLastErrorID;//sActErrorID
		Buffer_Act_Message[1].sModuleDescription:=sModuleDescription;

		//IF sActErrorID='000x000x999' THEN;
		//	Buffer_Act_Message[1].sErrorMessage:='General Error';	(*	Error description Not Found	*)
		//ELSE
			cFound:=0;
			FOR i:=1 TO C_Max_ErrorList DO
				IF ar_ErrorList[i,eErrID]=sActErrorID THEN
					iFound:=i;
					ar_ErrorActive[iFound]:=TRUE;
					cFound:=cFound+1;
				END_IF
			END_FOR
	
			IF cFound=1 THEN;
				Buffer_Act_Message[1].sErrorMessage:=ar_ErrorList[iFound,eErrMeassage];	(*	Error from the List	*)
				Buffer_Act_Message[1].sLevel:=ar_ErrorList[iFound,eErrLevel];	(*	Error Level from the List	*)
			ELSIF cFound=0 THEN; //(*	Error ID not Foud on the Error_List*)
				Buffer_Act_Message[1].sErrorMessage:='Error ID not found on the "Error_List"';	
				Buffer_Act_Message[1].sLevel:='Unknown';
			ELSIF cFound>1 THEN; //(*	More then one Errors Foud with the same  ID*)
				Buffer_Act_Message[1].sErrorMessage:='More then one error with the same ID  found on the "Error_list"';	
				Buffer_Act_Message[1].sLevel:='Unknown';
			END_IF
		//END_IF
		FUN_Write_Line_To_History();
	END_IF

END_FUNCTION_BLOCK

// ---- 00 Library/04-Messages/F_iFB_Num_sFB_Num.TcPOU
FUNCTION F_iFB_Num_sFB_Num : STRING(3)
VAR_INPUT
	iFB_Num: INT;
END_VAR
VAR
END_VAR

IF iFB_Num<10 THEN;
	F_iFB_Num_sFB_Num:=CONCAT(STR1:='00',STR2:=INT_TO_STRING(iFB_Num));
ELSIF iFB_Num<100 THEN;
	F_iFB_Num_sFB_Num:=CONCAT(STR1:='0',STR2:=INT_TO_STRING(iFB_Num));
ELSE;
	F_iFB_Num_sFB_Num:=CONCAT(STR1:='',STR2:=INT_TO_STRING(iFB_Num));
END_IF

END_FUNCTION

// ---- 00 Library/03 SFC/FB_SFC_Template.TcPOU
FUNCTION_BLOCK FB_SFC_Template EXTENDS FB_SFC_Cycle IMPLEMENTS ITF_FB_SFC_Cycle
VAR_INPUT
END_VAR
VAR_OUTPUT
END_VAR
VAR
END_VAR

m_Set_SFCFlags_Reference();
SUPER^();

ACTION act_Oper:
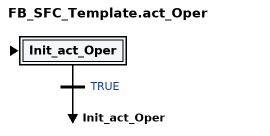
INITIAL_STEP Init_act_Oper:
END_STEP
TRANSITION FROM Init_act_Oper TO Init_act_Oper
    := TRUE;
END_TRANSITION
END_ACTION

METHOD m_Set_SFCFlags_Reference : BOOL
//Set reference to SFC flags

refSFC.SFCInit REF= SFCInit;
refSFC.SFCReset REF= SFCReset;
refSFC.SFCError REF= SFCError;
refSFC.SFCEnableLimit REF= SFCEnableLimit;
refSFC.SFCErrorStep REF= SFCErrorStep;
refSFC.SFCErrorPOU REF= SFCErrorPOU;
refSFC.SFCQuitError REF= SFCQuitError;
refSFC.SFCPause REF= SFCPause;
refSFC.SFCTrans REF= SFCTrans;
refSFC.SFCCurrentStep REF= SFCCurrentStep;
refSFC.SFCTip REF= SFCTip;
refSFC.SFCTipMode REF= SFCTipMode;

// Cycle handle for SFC
m_SFC_Handle();
END_METHOD

END_FUNCTION_BLOCK

// ---- 03 Project/00 -Initialise/prg_Initialise.TcPOU
PROGRAM prg_Initialise
VAR_INPUT
	ResumeSFC       : BOOL; 		(*	not automatic	*)
	//Added SFC Cycle handle Variables
	
	SFCInit             : BOOL;  //shachar
END_VAR

VAR


(* 8888888888888888   SFC   8888888888888888888888*)
	sCycleName	        : STRING;
	SFCCurrentStep      : STRING;
	SFCErrorPOU         : STRING;
	SFCErrorStep        : STRING;
	SFCError            : BOOL;
	SFCPause            : BOOL;
	
	SFCTipMode          : BOOL;
	SFCTip              : BOOL;
	SFCEnableLimit		: BOOL:=TRUE;
	// Reset Error
	SFCReset			: BOOL;
	ErrorSFC            : BOOL; 	(*	not automatic	*)

	ResetError          : BOOL; 	(*	not automatic	*)
	Last_SFCErrorStep   : STRING; 	(*	not automatic	*)
	//ErrorToPrint        : STRING; 	(*	not automatic	*)
	//Last_ErrorToPrint   : STRING; 	(*	not automatic	*)

 //   stSafety			:ST_BasicCycle;  //shachar
(* 8888888888888888   SFC   8888888888888888888888*)




	Pis             : INT;
	c_PisInitCheck  : INT;
	b_AllPisInitPos : BOOL;

	i               : INT;
	c_LatInitCheck  : INT;

	c_PisResetCleare: INT;

	k               : INT;

	bGeneralDone    : BOOL;
	bPistonDone     : BOOL;
	b_StationDone   : BOOL;
	bLoadConvDone   : BOOL;
	bUnloadConvDone : BOOL;
	bTableDone      : BOOL;
	bStackerDone    : BOOL;
    bManipulatorDone: BOOL;

	init_General    : BOOL;
	init_AllPiston  : BOOL;
	init_AllStation : BOOL;
	init_Table      : BOOL;
	init_LoadConv   : BOOL;
	init_UnloadConv : BOOL;
	init_Stacker    : BOOL;
	init_Manipulator: BOOL;

	bMessLoadInit   : BOOL;
	bMessUnloadInit : BOOL;
	
	sFB_ID          : STRING(4):='004';
	sFB_Num         : STRING(4):='000';
	sActErrorID     : STRING;
	//Added SFC Cycle handle Variables
	fb_SFC_Cycle		    : FB_SFC_Cycle;
	fbFormatString	    	: FB_FORMATSTRING;
	sFullErrorId		    : STRING(12);//sAAAxBBBxEEE
	bReset					: BOOL;

	bIntZoneOk: BOOL;
	bNotPrepare: BOOL;
	p_ManipReset: POINTER TO BOOL;
	p_PowerMotorOn: POINTER TO BOOL;
	p_SafetyStart: POINTER TO BOOL;
   // fbPowerMotorOn			:FB_PowerMotorOn;

	IndexOn: BOOL;
	LoadOn: BOOL;
	UnloadOn: BOOL;
	ManipOn: BOOL;
	p_PowerMotorPower: POINTER TO BOOL;
	p_PowerMotorOff: POINTER TO BOOL;
	iResumeCount: INT;
	iIndexCount: INT;
	iLoadCount: INT;
	iUnloadCount: INT;
	iManipCount: INT;
	p_ManipResume: POINTER TO BOOL;
END_VAR

VAR_IN_OUT
	stOperation	: ST_OperationButtons;	
END_VAR

act_General();
act_Piston();
act_GetErrorID();
fb_SFC_Cycle
( 
	sCycleName:= 'Initialize', 
	bSFCError:= SFCError, 
	sSFCCurrentStep:=SFCCurrentStep , 
	sSFCErrorStep:= SFCErrorStep, 
	sSFCErrorPOU:=SFCErrorPOU , 
	sActErrorID:=sFullErrorId,
	sFB_ModuleDescription:= fb_SFC_Cycle.sCycleName, 
	sLast_SFCErrorStep=>Last_SFCErrorStep , 
	bErrorSFC_Occured=> ErrorSFC, 
	//sErrorToPrint=>ErrorToPrint , 
	//sLast_ErrorToPrint=>Last_ErrorToPrint,
    bSFCInit=>SFCInit , 
	stOperation:= stOperation,
	bResumeSFC:=ResumeSFC , 
	bResetError:=ResetError , 
	bSFCPause:= SFCPause, 
	bResetCycle:=SFCReset
);



IF NOT bStateSafe	
OR init_AllPiston
THEN;
	bGeneralDone:=FALSE;
	bPistonDone:=FALSE;
	b_StationDone:=FALSE;
	bLoadConvDone:=FALSE;
	bUnloadConvDone:=FALSE;
	bTableDone:=FALSE;
	bStackerDone:=FALSE;
	bManipulatorDone:=FALSE;  //shachar
END_IF

ACTION act_General:
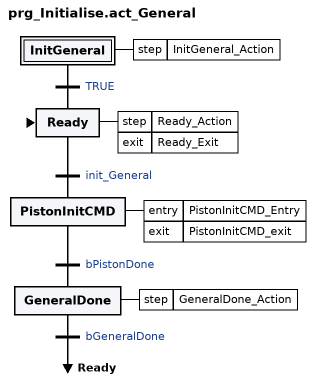
INITIAL_STEP InitGeneral:
    InitGeneral_Action(N);  // step action
END_STEP
TRANSITION FROM InitGeneral TO Ready
    := TRUE;
END_TRANSITION
STEP Ready:
    Ready_Action(N);  // step action
    Ready_Exit(P0);  // exit action
END_STEP
TRANSITION FROM Ready TO PistonInitCMD
    := init_General;
END_TRANSITION
STEP PistonInitCMD:  // min time t#2s
    PistonInitCMD_Entry(P1);  // entry action
    PistonInitCMD_exit(P0);  // exit action
END_STEP
TRANSITION FROM PistonInitCMD TO GeneralDone
    := bPistonDone;
END_TRANSITION
STEP GeneralDone:
    GeneralDone_Action(N);  // step action
END_STEP
TRANSITION FROM GeneralDone TO Ready
    := bGeneralDone;
END_TRANSITION
END_ACTION

ACTION act_GetErrorID:
IF ErrorSFC THEN;
	// Initialization
	IF    Last_SFCErrorStep='WatingForEmergencyOK' 			THEN sActErrorID:='001';
	ELSIF Last_SFCErrorStep='WatingForInterlockOK' 		    THEN sActErrorID:='002';
	ELSIF Last_SFCErrorStep='WatingForMotorsOK' 			THEN sActErrorID:='003';
	ELSIF Last_SFCErrorStep='CheckInitStationDone' 			THEN sActErrorID:='004';
	ELSIF Last_SFCErrorStep='Station_Initialization' 		THEN sActErrorID:='005';
	ELSIF Last_SFCErrorStep='Loader_Initialization' 		THEN sActErrorID:='006';
	ELSIF Last_SFCErrorStep='Unload_Station' 			    THEN sActErrorID:='007';
	ELSIF Last_SFCErrorStep='Measuring_Station' 			THEN sActErrorID:='008';
	ELSIF Last_SFCErrorStep='Gripper_Oriantation' 			THEN sActErrorID:='009';
	ELSIF Last_SFCErrorStep='Index_Homming' 			    THEN sActErrorID:='010';
	ELSIF Last_SFCErrorStep='PaletBypasCheck_1' 			THEN sActErrorID:='011';
	ELSIF Last_SFCErrorStep='PaletCheck_1' 			        THEN sActErrorID:='012';
	ELSIF Last_SFCErrorStep='Cover_Station' 			    THEN sActErrorID:='023';	
	ELSE;
		 sActErrorID:='999';
	END_IF
//ELSIF bWarning THEN;
	// Leave the warning message to print
ELSE;
		 sActErrorID:='000';
END_IF
//*** Error Format ***
fbFormatString(
	sFormat:= '%.3sx%.3sx%.3s', 
	arg1:= F_STRINGEx(sFB_ID), 
	arg2:= F_STRINGEx(sFB_Num), 
	arg3:= F_STRINGEx(sActErrorID), 
	sOut=>sFullErrorId );
	
//(*Clean Last ErrID*)IF NOT SFCPause THEN	sFullErrorId:='';END_IF
END_ACTION

ACTION act_Piston:
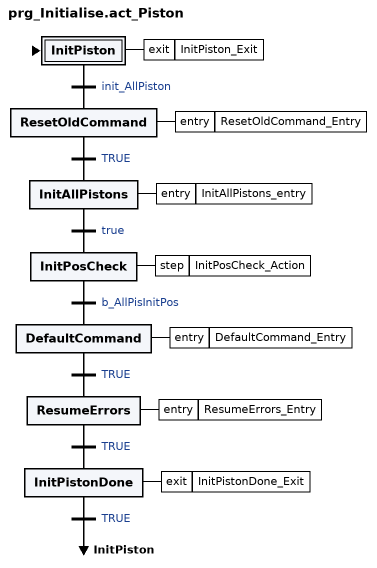
INITIAL_STEP InitPiston:
    InitPiston_Exit(P0);  // exit action
END_STEP
TRANSITION FROM InitPiston TO ResetOldCommand
    := init_AllPiston;
END_TRANSITION
STEP ResetOldCommand:  // min time T#0.1S
    ResetOldCommand_Entry(P1);  // entry action
END_STEP
TRANSITION FROM ResetOldCommand TO InitAllPistons
    := TRUE;
END_TRANSITION
STEP InitAllPistons:  // min time t#1s
    InitAllPistons_entry(P1);  // entry action
END_STEP
TRANSITION FROM InitAllPistons TO InitPosCheck
    := true;
END_TRANSITION
STEP InitPosCheck:
    InitPosCheck_Action(N);  // step action
END_STEP
TRANSITION FROM InitPosCheck TO DefaultCommand
    := b_AllPisInitPos;
END_TRANSITION
STEP DefaultCommand:  // min time T#0.2S
    DefaultCommand_Entry(P1);  // entry action
END_STEP
TRANSITION FROM DefaultCommand TO ResumeErrors
    := TRUE;
END_TRANSITION
STEP ResumeErrors:  // min time T#0.2S
    ResumeErrors_Entry(P1);  // entry action
END_STEP
TRANSITION FROM ResumeErrors TO InitPistonDone
    := TRUE;
END_TRANSITION
STEP InitPistonDone:
    InitPistonDone_Exit(P0);  // exit action
END_STEP
TRANSITION FROM InitPistonDone TO InitPiston
    := TRUE;
END_TRANSITION
END_ACTION

ACTION DefaultCommand_Entry:
	(*FOR Pis:=1 TO 24 BY 1 DO
		db_Lat[Pis].req_DefaultPos:=TRUE;
	END_FOR*)
	
	FOR Pis:=1 TO C_Max_Pistons BY 1 DO
		IF stPis[Pis].b_PistonActive THEN;
			stPis[Pis].req_Init:=TRUE;
		END_IF		
	END_FOR
END_ACTION

ACTION GeneralDone_Action:
init_General:=FALSE;
bGeneralDone:=TRUE;
END_ACTION

ACTION InitAllPistons_entry:
prg_Pistons.bInitAllPiston:=TRUE;
END_ACTION

ACTION InitGeneral_Action:
SFCReset:=FALSE;

init_AllPiston   :=FALSE;
END_ACTION

ACTION InitPiston_Exit:
	b_AllPisInitPos:=FALSE;
	bPistonDone:=FALSE;
END_ACTION

ACTION InitPistonDone_Exit:
	init_AllPiston:=FALSE;
	bPistonDone:=TRUE;
END_ACTION

ACTION InitPosCheck_Action:
			c_PisInitCheck:=0;
	FOR Pis:=1 TO C_Max_Pistons BY 1 DO
		IF fb_Pis[Pis].SFCCurrentStep<>'Ready' AND fb_Pis[Pis].SFCCurrentStep<>''THEN
			c_PisInitCheck:=c_PisInitCheck+1;
		END_IF
	END_FOR

			c_PisResetCleare:=0;
	FOR Pis:=1 TO C_Max_Pistons BY 1 DO
		IF stPis[Pis].b_Reset THEN
			c_PisResetCleare:=c_PisResetCleare+1;
		END_IF
	END_FOR

	(*		c_LatInitCheck:=0;
	FOR Pis:=1 TO 24 BY 1 DO
		IF fb_Lat[Pis].SFCCurrentStep<>'Ready' AND fb_Lat[Pis].SFCCurrentStep<>'' THEN
			c_LatInitCheck:=c_LatInitCheck+1;
		END_IF
	END_FOR*)


		IF 	c_PisInitCheck=0  AND c_LatInitCheck=0 (*AND 	c_PisResetCleare=0*) THEN
			b_AllPisInitPos:=TRUE;
		ELSE
			b_AllPisInitPos:=FALSE;
		END_IF
END_ACTION

ACTION PistonInitCMD_Entry:
init_AllPiston:=TRUE;
END_ACTION

ACTION PistonInitCMD_exit:
Global_Variables.ResumeAll :=TRUE;
END_ACTION

ACTION Ready_Action:
IF TRUE
AND	bPistonDone
(*AND	b_StationDone
AND	bLoadConvDone
AND	bUnloadConvDone
AND	bTableDone
AND (bManipulatorDone OR NOT b_ManipulatorExist)
AND	(bStackerDone OR NOT b_StackerExist)*)
THEN
	bGeneralDone:=TRUE;

ELSE
	bGeneralDone:=FALSE;
END_IF
END_ACTION

ACTION Ready_Exit:
bGeneralDone:=FALSE;
bPistonDone:=FALSE;
b_StationDone:=FALSE;
bLoadConvDone:=FALSE;
bUnloadConvDone:=FALSE;
bTableDone:=FALSE;
bStackerDone:=FALSE;

bManipulatorDone:=FALSE; //shachar
iResumeCount:=0;
END_ACTION

ACTION ResetOldCommand_Entry:
	(*FOR Pis:=1 TO 24 BY 1 DO
		db_Lat[Pis].req_Reset:=TRUE;
	END_FOR*)
	FOR Pis:=1 TO C_Max_Pistons BY 1 DO
		stPis[Pis].b_Reset:=TRUE;
	END_FOR
END_ACTION

ACTION ResumeErrors_Entry:
	(*FOR Pis:=1 TO 24 BY 1 DO
		db_Lat[Pis].req_Resume:=TRUE;
	END_FOR*)
	FOR Pis:=1 TO C_Max_Pistons BY 1 DO
		stPis[Pis].b_Resume:=TRUE;
	END_FOR
END_ACTION

END_PROGRAM

// ---- 03 Project/15 Production Recipes/FB_ProdRecipe_Manage.TcPOU
FUNCTION_BLOCK FB_ProdRecipe_Manage
VAR_INPUT
END_VAR
VAR_OUTPUT
END_VAR
VAR
	stProdParam_HMI: ST_Production_Parameter;

	bReInit: BOOL;
END_VAR

IF bReInit THEN;
	FB_INIT(bInCopyCode:=FALSE,bInitRetains:=FALSE);
	bReInit:=FALSE;
	//FB_INIT.bInitRetains:=TRUE;
END_IF
mPercentage_Calculation();
mGet_Recipe_list();

g_Prod.dtProdTimeMin:=dtRealTime-T#2H;
g_Prod.dtProdTimeMax:=dtRealTime+T#7D;

METHOD FB_INIT : BOOL
VAR_INPUT
END_VAR
VAR_INPUT
    bInitRetains : BOOL; // TRUE if the FB is being initialized after a warm restart
    bInCopyCode : BOOL;  // TRUE if the FB is being initialized in copy code
END_VAR
VAR
	i: INT;
	k: INT;
END_VAR
FOR i:=0 TO g_Prod.cMax_Prod_Recipe DO
	
	g_Prod.arrRecipeMarinade[i].prodType:=E_Prod_Type.Marinade;
	g_Prod.arrRecipeColor[i].prodType:=E_Prod_Type.Color;
	
	g_Prod.arrRecipeMarinade[i].arr_Component[1].sDescription:='Water';
	g_Prod.arrRecipeColor[i].arr_Component[1].sDescription:='Water';
	
	g_Prod.arrRecipeMarinade[i].arr_Component[1].eIngredientType:=E_Ingredient_type.eWater;
	g_Prod.arrRecipeColor[i].arr_Component[1].eIngredientType:=E_Ingredient_type.eWater;

	FOR k:=2 TO g_Prod.cMaxCompInProduct-1 DO
		//g_Prod.arrRecipeMarinade[i].arr_Component[k].sDescription:='Powder';
		//g_Prod.arrRecipeColor[i].arr_Component[k].sDescription:='Powder';
		
		g_Prod.arrRecipeMarinade[i].arr_Component[k].eIngredientType:=E_Ingredient_type.ePowder;
		g_Prod.arrRecipeColor[i].arr_Component[k].eIngredientType:=E_Ingredient_type.ePowder;		
	END_FOR
	
	
	
	g_Prod.arrRecipeMarinade[i].arr_Component[10].sDescription:='Oil';
	g_Prod.arrRecipeColor[i].arr_Component[10].sDescription:='Oil';
	
	g_Prod.arrRecipeMarinade[i].arr_Component[10].eIngredientType:=E_Ingredient_type.eOil;
	g_Prod.arrRecipeColor[i].arr_Component[10].eIngredientType:=E_Ingredient_type.eOil;	

END_FOR
END_METHOD

METHOD mGet_Recipe_list : BOOL
VAR_INPUT
END_VAR

VAR
	i: INT;
END_VAR
FOR i:=1 TO g_Prod.cMax_Prod_Recipe DO
	g_Prod.listRecipe_Marinade[i]:=g_Prod.arrRecipeMarinade[i].Description;
	g_Prod.listRecipe_Color[i]:=g_Prod.arrRecipeColor[i].Description;
	
	
END_FOR
END_METHOD

METHOD mPercentage_Calculation : BOOL
VAR_INPUT
END_VAR

VAR
	i: INT;
	tempPercentage_M: REAL;
	tempPercentage_C: REAL;
	k: INT;
END_VAR

FOR i:=1 TO g_Prod.cMax_Prod_Recipe DO
	tempPercentage_M:=0;
	tempPercentage_C:=0;	
	FOR k:=2 TO g_Prod.cMaxCompInProduct DO
		tempPercentage_M:=tempPercentage_M + g_Prod.arrRecipeMarinade[i].arr_Component[k].rWeightPercentage;
		tempPercentage_C:=tempPercentage_C + g_Prod.arrRecipeColor[i].arr_Component[k].rWeightPercentage;
	END_FOR
	g_Prod.arrRecipeMarinade[i].arr_Component[1].rWeightPercentage:=100-tempPercentage_M;
	g_Prod.arrRecipeColor[i].arr_Component[1].rWeightPercentage:=100-tempPercentage_C;
END_FOR
END_METHOD

END_FUNCTION_BLOCK

// ---- 00 Library/00-General/CheckBounds.TcPOU
FUNCTION CheckBounds : DINT
VAR_INPUT
	index, lower, upper : DINT;
END_VAR
VAR
END_VAR

IF index<lower THEN
	CheckBounds := lower;
	Errors:=Errors+1;
ELSIF index>upper THEN
	CheckBounds := upper;
	Errors:=Errors+1;
ELSE
	CheckBounds := index;
END_IF

END_FUNCTION

// ---- 00 Library/00-General/TimeAndDate/FUN_DeltaTime.TcPOU
FUNCTION FUN_DeltaTime : STRING
VAR_INPUT
    //stSystemTime : TimeStruct;
    stStartTime  : TimeStruct;	
END_VAR
VAR
    dtSystemTime : DT;
    dtStartTime  : DT;
    deltaTime    : TIME;
    hours        : INT;
    minutes      : INT;
    milliseconds : INT;
    sDeltaTime   : STRING;	
END_VAR

// Convert TimeStruct to DT
dtSystemTime := SYSTEMTIME_TO_DT(stSystemTime);
dtStartTime  := SYSTEMTIME_TO_DT(stStartTime);

// Calculate the delta time
deltaTime := TO_TIME(dtSystemTime - dtStartTime);

// Extract hours, minutes, and milliseconds
hours := INT_TO_DINT(deltaTime / T#1H);
minutes := INT_TO_DINT((deltaTime MOD T#1H) / T#1M);
milliseconds := INT_TO_DINT((deltaTime MOD T#1M) / T#1MS);

// Format the string
sDeltaTime := CONCAT(CONCAT(CONCAT(CONCAT(INT_TO_STRING(hours), ':'), INT_TO_STRING(minutes)), ':'), INT_TO_STRING(milliseconds));

FUN_DeltaTime := sDeltaTime;

END_FUNCTION

// ---- 00 Library/04 Recipe/OLD/prg_RecipeManager.TcPOU
PROGRAM prg_RecipeManager
VAR
	fbRecipe: RecipeManCommands;
	LastError: DWORD;
	LastInfo: InfoValues;

	bCheckError: BOOL;
	bResetError: BOOL;
	bInit: BOOL;
END_VAR


IF bCheckError THEN;
	//bCheckError:=FALSE;
	LastError:=fbRecipe.GetLastError();
	LastInfo:=fbRecipe.GetLastInfo();
END_IF

IF bResetError THEN;
	bResetError:=FALSE;
	LastError:=fbRecipe.ResetLastError();
	LastError:=fbRecipe.ReloadRecipes(RecipeDefinitionName:='');
	
END_IF

IF bInit THEN;
	bInit:=FALSE;
	LastError:=fbRecipe.ResetLastInfo();
END_IF

END_PROGRAM

// ---- 00 Library/04-Messages/FB_PrintErrMessageByID_ST_Cycle.TcPOU
FUNCTION_BLOCK FB_PrintErrMessageByID_ST_Cycle
VAR_INPUT
	pstCycle			:POINTER TO ST_BasicCycle;
	sActErrorID			: STRING;
	ErrorToPrint		: STRING;
	iFB_Num				: INT:=0;
	sFB_ModuleDescription	:STRING(30):='';
	bResumeAll		: BOOL;
END_VAR
VAR_OUTPUT
END_VAR
VAR
	cFound				: INT;
	i					: INT;
	iFound				: INT;
	//r_trigPrintMessage	: R_TRIG;
	bNewMeasege			: BOOL;
	sActErrorID_AA		: STRING;
	iErrorID_Flag		: INT;
	sAA					: STRING;
	sActErrorID_Message	: STRING;
	iAAPos				: INT;
	rtrig1				: R_TRIG;
	
	sLastErrorID: STRING;
	j: INT;
END_VAR


IF pstCycle^.bFault THEN
	IF sActErrorID<>'000x000x000'  AND sActErrorID<>'' THEN //to print or not to print the massage???
		sLastErrorID:=sActErrorID;
		bNewMeasege:=TRUE;
		FOR i:=1 TO 100 DO
			IF Buffer_Act_Message[i].sErrID=sActErrorID THEN;
				IF Buffer_Act_Message[i].sModuleDescription = sFB_ModuleDescription THEN
					bNewMeasege:=FALSE;
					EXIT;
				END_IF
			END_IF
		END_FOR
	ELSE
		bNewMeasege:=FALSE;
	END_IF
	
	IF bNewMeasege AND NOT bResumeAll THEN;
		FOR i:=100 TO 2 BY -1 DO
			Buffer_Act_Message[i].sDateTime:=Buffer_Act_Message[i-1].sDateTime;
			Buffer_Act_Message[i].sErrID:=Buffer_Act_Message[i-1].sErrID;
			Buffer_Act_Message[i].sErrorMessage:=Buffer_Act_Message[i-1].sErrorMessage;
			Buffer_Act_Message[i].sLevel:=Buffer_Act_Message[i-1].sLevel;
			Buffer_Act_Message[i].sModuleDescription:=Buffer_Act_Message[i-1].sModuleDescription;
		END_FOR
		
		Buffer_Act_Message[1].sDateTime:=prg_RealClock.sRealTime_Date;
		Buffer_Act_Message[1].sErrID:=sActErrorID;
		Buffer_Act_Message[1].sModuleDescription:=sFB_ModuleDescription;

		IF sActErrorID='000x000x999' THEN;
			Buffer_Act_Message[1].sErrorMessage:=CONCAT('Cycle message: ',ErrorToPrint);
		ELSE
			cFound:=0;
			FOR i:=1 TO C_Max_ErrorList DO
				IF ar_ErrorList[i,eErrID]=sActErrorID THEN
					iFound:=i;
					ar_ErrorActive[iFound]:=TRUE;
					cFound:=cFound+1;
				END_IF
			END_FOR
	
			IF cFound=1 THEN;
				Buffer_Act_Message[1].sErrorMessage:=ar_ErrorList[iFound,eErrMeassage];	(*	Error from the List	*)
				pstCycle^.sFailedMessage := Buffer_Act_Message[1].sErrorMessage;
				Buffer_Act_Message[1].sLevel:=ar_ErrorList[iFound,eErrLevel];	(*	Error Level from the List	*)
			ELSIF cFound=0 THEN; //(*	Error ID not Foud on the List	*)
				//Buffer_Act_Message[1].sErrorMessage:='Error ID not found on the "Error List"';
				Buffer_Act_Message[1].sErrorMessage:=CONCAT('Cycle message[1]: ',ErrorToPrint);
				Buffer_Act_Message[1].sLevel:='Error';
			ELSIF cFound>1 THEN; //(*	More then one Errors Foud with the same  ID		*)
				//Buffer_Act_Message[1].sErrorMessage:='More then one error with the same ID  found on the "Error list"';
				Buffer_Act_Message[1].sErrorMessage:=CONCAT('Cycle message[2]: ',ErrorToPrint);
				Buffer_Act_Message[1].sLevel:='Error';
			END_IF
		END_IF
		FUN_Write_Line_To_History();
	END_IF
	
	
	IF bResumeAll THEN
		sActErrorID:='';
	END_IF
	
END_IF

(*
//for delete message if no fault
rtrig1(CLK:= NOT pstCycle^.bFault, Q=> );
IF rtrig1.Q THEN  // if cycle not in pause
	FOR i:= 2 TO 100 DO //loop for search 
		IF Buffer_Act_Message[i-1].sErrID = sLastErrorID THEN // search if last error id = buffer which it error table.
			FOR j:= i TO 100 DO //if found message id then delete it.
				Buffer_Act_Message[j-1]:=Buffer_Act_Message[j];//delete
			END_FOR
		END_IF
	END_FOR
END_IF
*)

END_FUNCTION_BLOCK

// ---- 00 Library/07 Errors/FB_Error_Handle.TcPOU
FUNCTION_BLOCK FB_Error_Handle
VAR_INPUT
	bError: BOOL;
	sErrID: STRING;
END_VAR
VAR_OUTPUT
END_VAR
VAR
	fbFormat: FB_FormatString;
END_VAR
VAR_IN_OUT
	error_code: STRING;

END_VAR



IF bError 
AND error_code=''
THEN;
	error_code:=sErrID;
END_IF

IF NOT bError 
AND error_code=sErrID
THEN;
	error_code:='';
END_IF

METHOD m_GetAxisErr : STRING(4)
VAR_INPUT
	stDevErr_H				: ST_DeviceErrorHandeling;
END_VAR
VAR_OUTPUT
	sMessage: STRING;
END_VAR

VAR
	ErrID_xx: STRING(2);
END_VAR
IF bError 
AND error_code=''
THEN;
	fbFormat(sFormat:='%0.2d' ,arg1:=F_INT(stDevErr_H.iObjectID),sOut=>ErrID_xx);
	m_GetAxisErr:=CONCAT('23',ErrID_xx);
	sMessage:=stDevErr_H.sObjectName;
ELSE;
	m_GetAxisErr:='';
END_IF
END_METHOD

METHOD m_GetPistonErr : STRING(4)
VAR_INPUT
	stDevErr_H				: ST_DeviceErrorHandeling;
END_VAR
VAR_OUTPUT
	sMessage: STRING;
END_VAR

VAR
	ErrID_xx: STRING(2);
END_VAR
IF bError 
AND error_code=''
THEN;
	fbFormat(sFormat:='%0.2d' ,arg1:=F_INT(stDevErr_H.iObjectID),sOut=>ErrID_xx);
	m_GetPistonErr:=CONCAT('22',ErrID_xx);
	sMessage:=stDevErr_H.sObjectName;
ELSE;
	m_GetPistonErr:='';
END_IF
END_METHOD

END_FUNCTION_BLOCK

// ---- 00 Library/10 Utils/DutyCycle/FB_DutyCycle.TcPOU
FUNCTION_BLOCK FB_DutyCycle
VAR_INPUT
	bEnable		: BOOL;
	fBaseTime	: REAL:=5.0; // [sec] min>0
	fOn_Duty	: REAL:=10.0; //min =0, max=100
END_VAR
VAR_OUTPUT
	bOut: BOOL;
END_VAR
VAR
	tBaseTime: TIME;
	ton_OnDuty: TON;
	fOnTime: REAL;
	tOnTime: TIME;
END_VAR


tBaseTime:=REAL_TO_TIME(fBaseTime*1000);
ton_OnDuty(PT:=tBaseTime,IN:=NOT ton_OnDuty.Q AND bEnable);

IF fOn_Duty<0 THEN;
	fOn_Duty:=0;
ELSIF fOn_Duty>100 THEN;
	fOn_Duty:=1000;
END_IF
	
fOnTime:=fBaseTime*fOn_Duty/100.0;
tOnTime:=REAL_TO_TIME(fOnTime*1000);

IF bEnable THEN;
	IF fOn_Duty<=0 THEN;
		bOut:=FALSE;
	ELSIF fOn_Duty>=100 THEN;
		bOut:=TRUE;
	ELSE;
		IF ton_OnDuty.ET<tOnTime THEN;
			bOut:=TRUE;
		ELSE
			bOut:=FALSE;
		END_IF		
	END_IF	
ELSE;
	bOut:=FALSE;
END_IF

END_FUNCTION_BLOCK

// ---- 00 Library/10 Utils/fun_LrealToString.TcPOU
FUNCTION fun_LrealToString : STRING
VAR_INPUT
	iDigits	: INT:=2;
	fVar	: LREAL;
END_VAR
VAR
	iDigitsLocal: INT;

	fTemp: LREAL;
	fMult: LREAL;
	
	fbFormat: FB_FormatString;	

END_VAR

IF iDigits<0 THEN;
	iDigitsLocal:=0;
ELSIF iDigits>6 THEN;
	iDigitsLocal:=6; 
ELSE
	iDigitsLocal:=iDigits;	
END_IF

// this vertion solve the case then the result is 2.0-e2 instade of 0.02
CASE iDigitsLocal OF
	0:;fbFormat(sFormat:='%.0f' ,arg1:=F_LREAL(fVar),sOut=>fun_LrealToString);
	1:;fbFormat(sFormat:='%.1f' ,arg1:=F_LREAL(fVar),sOut=>fun_LrealToString);
	2:;fbFormat(sFormat:='%.2f' ,arg1:=F_LREAL(fVar),sOut=>fun_LrealToString);
	3:;fbFormat(sFormat:='%.3f' ,arg1:=F_LREAL(fVar),sOut=>fun_LrealToString);
	4:;fbFormat(sFormat:='%.4f' ,arg1:=F_LREAL(fVar),sOut=>fun_LrealToString);
	5:;fbFormat(sFormat:='%.5f' ,arg1:=F_LREAL(fVar),sOut=>fun_LrealToString);
	6:;fbFormat(sFormat:='%.6f' ,arg1:=F_LREAL(fVar),sOut=>fun_LrealToString);
END_CASE

(* OLD Version
CASE iDigitsLocal OF
	0:;fMult:=1;
	1:;fMult:=10;
	2:;fMult:=100;
	3:;fMult:=1000;
	4:;fMult:=10000;
	5:;fMult:=100000;
	6:;fMult:=1000000;
END_CASE

fTemp:=TRUNC(fVar*fMult);
IF iDigitsLocal=0 THEN;
	fun_LrealToString:=DINT_TO_STRING(TRUNC(fVar));
ELSE;
	fun_LrealToString:=LREAL_TO_STRING(fTemp/fMult);	
END_IF
*)

END_FUNCTION

// ---- 00 Library/10 Utils/F_TimeRatio.TcPOU
FUNCTION F_TimeRatio : INT
VAR_INPUT
	t1: TIME;
	t2: TIME;

END_VAR
VAR
	udi_t1: UDINT;
	udi_t2: UDINT;

	ratio: REAL;
END_VAR


udi_t1:=TIME_TO_UDINT(t1);
udi_t2:=TIME_TO_UDINT(t2);

IF udi_t2>0 THEN;
	ratio:=udi_t1/udi_t2;
END_IF

END_FUNCTION

// ---- 01 Instance/04-Messages/Prg_Filter_Messages.TcPOU
PROGRAM Prg_Filter_Messages
VAR
	sSearchMessage		: STRING;
	i					: INT;
	d					: INT;
	stFilter			: stMessageFormat;
	stLastFilter		: stMessageFormat;
	T1					: TON;
	bFilter				: BOOL;
END_VAR


IF stFilter.sErrID<>stLastFilter.sErrID
OR  stFilter.sLevel <>stLastFilter.sLevel
OR  stFilter.sModuleDescription <>stLastFilter.sModuleDescription
OR  stFilter.sErrorMessage<>stLastFilter.sErrorMessage THEN

	FOR i:=1000 TO 1 BY -1 DO
		Buffer_Search_Messages[i].sDateTime:='';
		Buffer_Search_Messages[i].sErrID:='';
		Buffer_Search_Messages[i].sErrorMessage:='';
		Buffer_Search_Messages[i].sLevel:='';
		Buffer_Search_Messages[i].sModuleDescription:='';
	END_FOR
	bFilter:=TRUE;
ELSE
	bFilter:=FALSE;
END_IF




T1(IN:=bFilter , PT:=T#300MS , Q=> , ET=> );
IF T1.Q THEN
	d:=2;
	FOR i:=1 TO 1000 DO
			IF (Buffer_Act_History[i].sErrID=stFilter.sErrID OR stFilter.sErrID='')
			AND (Buffer_Act_History[i].sLevel=stFilter.sLevel OR stFilter.sLevel='')
			AND (Buffer_Act_History[i].sErrorMessage=stFilter.sErrorMessage OR stFilter.sErrorMessage='')
			AND (Buffer_Act_History[i].sModuleDescription=stFilter.sModuleDescription OR stFilter.sModuleDescription='')THEN
				Buffer_Search_Messages[d]:=Buffer_Act_History[i];
				d:=d+1;
			END_IF
	END_FOR
	
	
ELSE

FOR i:=1000 TO 2 BY -1 DO
	Buffer_Search_Messages[i]:=Buffer_Act_History[i-1];
END_FOR

END_IF

END_PROGRAM

// ---- 01 Instance/07-Mode/prg_HMI_OperationLock.TcPOU
PROGRAM prg_HMI_OperationLock
VAR
	b_LockIndex: BOOL;
	b_LockLoad: BOOL;
	b_LockUnload: BOOL;
	b_LockManip: BOOL;
END_VAR

IF stModeMain.iActMode= 2 AND prg_User.actUser< 3 THEN
   b_LockIndex := TRUE;
ELSE
   b_LockIndex := FALSE;
END_IF

END_PROGRAM

// ---- 03 Project/13 Weight control/FB_FillingMarinade.TcPOU
FUNCTION_BLOCK FB_FillingMarinade
VAR_INPUT
	iFillAmoungKg		: UINT;
	rActWeight			: REAL;
	bStop				: BOOL;
END_VAR
VAR_OUTPUT
	bFillingBusy		: BOOL;
	bFillingDone		: BOOL;
END_VAR
VAR_IN_OUT
	bFillRequest		: BOOL;
	fbFiliingPump		: FB_Pump;
	bPistonOpen			: BOOL;
	bPistonClose		: BOOL;
END_VAR
VAR
	trigStop			: R_TRIG;
	rHighVelocity		: REAL:=200;
	rMidVelocity		: REAL:=100;
	rLowVelocity		: REAL:=10;
END_VAR

actFillComponent();

trigStop(Clk:= bStop);
IF SFCReset THEN
	SFCReset:=FALSE;
END_IF
IF trigStop.Q THEN
	bFillRequest:=FALSE;
	SFCReset:=TRUE;
END_IF

ACTION actFillComponent:
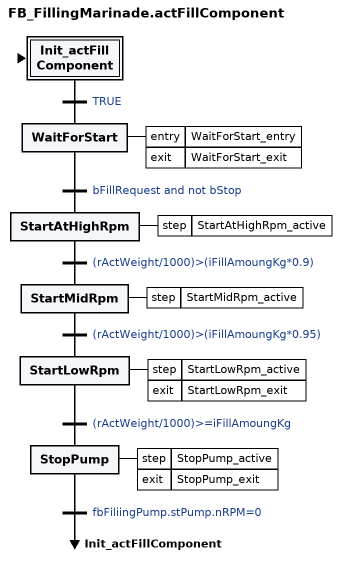
INITIAL_STEP Init_actFillComponent:
END_STEP
TRANSITION FROM Init_actFillComponent TO WaitForStart
    := TRUE;
END_TRANSITION
STEP WaitForStart:
    WaitForStart_entry(P1);  // entry action
    WaitForStart_exit(P0);  // exit action
END_STEP
TRANSITION FROM WaitForStart TO StartAtHighRpm
    := bFillRequest and not bStop;
END_TRANSITION
STEP StartAtHighRpm:
    StartAtHighRpm_active(N);  // step action
END_STEP
TRANSITION FROM StartAtHighRpm TO StartMidRpm
    := (rActWeight/1000)>(iFillAmoungKg*0.9);
END_TRANSITION
STEP StartMidRpm:
    StartMidRpm_active(N);  // step action
END_STEP
TRANSITION FROM StartMidRpm TO StartLowRpm
    := (rActWeight/1000)>(iFillAmoungKg*0.95);
END_TRANSITION
STEP StartLowRpm:
    StartLowRpm_active(N);  // step action
    StartLowRpm_exit(P0);  // exit action
END_STEP
TRANSITION FROM StartLowRpm TO StopPump
    := (rActWeight/1000)>=iFillAmoungKg;
END_TRANSITION
STEP StopPump:
    StopPump_active(N);  // step action
    StopPump_exit(P0);  // exit action
END_STEP
TRANSITION FROM StopPump TO Init_actFillComponent
    := fbFiliingPump.stPump.nRPM=0;
END_TRANSITION
END_ACTION

ACTION StartAtHighRpm_active:
fbFiliingPump.m_Run(RPM:=rHighVelocity);
END_ACTION

ACTION StartLowRpm_active:
fbFiliingPump.m_Run(RPM:=rMidVelocity);
END_ACTION

ACTION StartLowRpm_exit:
bPistonOpen:=FALSE;
bPistonClose:=TRUE;
END_ACTION

ACTION StartMidRpm_active:
fbFiliingPump.m_Run(RPM:=rMidVelocity);
END_ACTION

ACTION StopPump_active:
fbFiliingPump.m_Stop();
END_ACTION

ACTION StopPump_exit:
bFillingBusy:=FALSE;		
bFillingDone:=TRUE;
END_ACTION

ACTION WaitForStart_entry:
fbFiliingPump.m_Stop();
bPistonOpen:=FALSE;
bPistonClose:=TRUE;
END_ACTION

ACTION WaitForStart_exit:
bFillingBusy:=TRUE;		
bFillingDone:=FALSE;
bPistonOpen:=TRUE;
bPistonClose:=FALSE;
END_ACTION

END_FUNCTION_BLOCK

// ---- 03 Project/13 Weight control/Production/FB_SetProductionParams.TcPOU
FUNCTION_BLOCK FB_SetProductionParams
VAR_INPUT
END_VAR
VAR_OUTPUT
	rCompActualWeight	: REAL;
	iCoun: INT;
	i:INT;
END_VAR
VAR_IN_OUT
	stProdParams		: ST_ProdParams;
	stTriBlender		: ST_TriBlender;
	bTankInProduction	: BOOL;
END_VAR
VAR_INPUT
	iActualWaterAmount	: UINT;
END_VAR


rCompActualWeight:=(TO_REAL(iActualWaterAmount)/100)*stProdParams.arrComponents[i].rCompWeightFor100L;

ACTION act_SetProdVal:

END_ACTION

END_FUNCTION_BLOCK

// ---- 03 Project/13 Weight control/TriBlender/POUs/prg_TriBlender.TcPOU
PROGRAM prg_TriBlender
VAR
	enumCurrentState	: ENUM_CurrentState;
	FB_SetProductionParams:FB_SetProductionParams;
//stTriBlender		: ST_TriBlender;
	
	sStateDescription		: STRING;
	sStateInstructions		: STRING;
	iCirculationTimeLeft	: UINT;
	bContinue				: BOOL;
	iCurrentMixingComponent	: INT;
	
	tonStageCirculation		: TON;
	
	///For Visu
	bDisableTime			: BOOL;
	bDisableAmount			: BOOL;
	bDisableName			: BOOL;
	bDisableButton			: BOOL;
	wButtonColor			: DWORD;
	
	trig_JumpToCirScreen	: R_TRIG;

	i						: INT;
	bTesting: BOOL;
END_VAR
VAR_IN_OUT
	stTriblender			: ST_TriBlender;
	fb_TriBlenderPump		: FB_Pump;
END_VAR
VAR_INPUT
	arrComponents	: ARRAY [0..g_Prod.cMaxCompInProduct-1] OF ST_Component;
END_VAR

trig_JumpToCirScreen(CLK:= stTriblender.bStartDisolving);

IF trig_JumpToCirScreen.Q THEN
	VisuElems.CurrentVisu:= 'Main';	
END_IF

Init_act_MixingStates();

stTriblender.bPumpOnFdbk:= fb_TriBlenderPump.bRun;

FB_SetProductionParams(stProdParams:=g_Data.arr_ProdTank[0],bTankInProduction:=bTesting,iActualWaterAmount:=100,stTriBlender:=g_Data.stTriBlender);

ACTION CheckIfLast_entry:
bDisableButton:=FALSE;

fb_TriBlenderPump.m_Stop();
bContinue:=FALSE;
END_ACTION

ACTION FlowOrPressureError_entry:
stTriblender.bError:=TRUE;
stTriblender.sErrorDescription:='Pressure or flow error';
VisuElems.CurrentVisu:= 'StartVisu';
END_ACTION

ACTION Init_act_MixingStates:
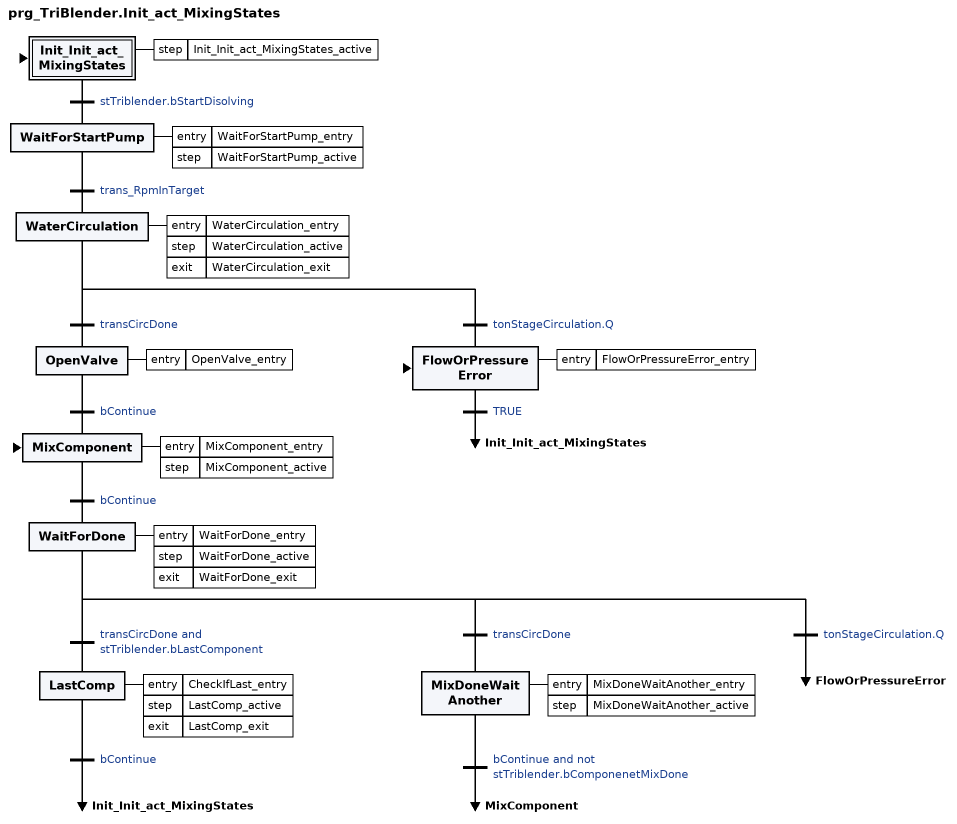
INITIAL_STEP Init_Init_act_MixingStates:
    Init_Init_act_MixingStates_active(N);  // step action
END_STEP
TRANSITION FROM Init_Init_act_MixingStates TO WaitForStartPump
    := stTriblender.bStartDisolving;
END_TRANSITION
STEP WaitForStartPump:
    WaitForStartPump_entry(P1);  // entry action
    WaitForStartPump_active(N);  // step action
END_STEP
TRANSITION FROM WaitForStartPump TO WaterCirculation
    := trans_RpmInTarget;
END_TRANSITION
STEP WaterCirculation:
    WaterCirculation_entry(P1);  // entry action
    WaterCirculation_active(N);  // step action
    WaterCirculation_exit(P0);  // exit action
END_STEP
TRANSITION FROM WaterCirculation TO OpenValve
    := transCircDone;
END_TRANSITION
TRANSITION FROM WaterCirculation TO FlowOrPressureError
    := tonStageCirculation.Q;
END_TRANSITION
STEP FlowOrPressureError:
    FlowOrPressureError_entry(P1);  // entry action
END_STEP
TRANSITION FROM FlowOrPressureError TO Init_Init_act_MixingStates
    := TRUE;
END_TRANSITION
STEP OpenValve:
    OpenValve_entry(P1);  // entry action
END_STEP
TRANSITION FROM OpenValve TO MixComponent
    := bContinue;
END_TRANSITION
STEP MixComponent:
    MixComponent_entry(P1);  // entry action
    MixComponent_active(N);  // step action
END_STEP
TRANSITION FROM MixComponent TO WaitForDone
    := bContinue;
END_TRANSITION
STEP WaitForDone:
    WaitForDone_entry(P1);  // entry action
    WaitForDone_active(N);  // step action
    WaitForDone_exit(P0);  // exit action
END_STEP
TRANSITION FROM WaitForDone TO LastComp
    := transCircDone and stTriblender.bLastComponent;
END_TRANSITION
TRANSITION FROM WaitForDone TO MixDoneWaitAnother
    := transCircDone;
END_TRANSITION
TRANSITION FROM WaitForDone TO FlowOrPressureError
    := tonStageCirculation.Q;
END_TRANSITION
STEP MixDoneWaitAnother:
    MixDoneWaitAnother_entry(P1);  // entry action
    MixDoneWaitAnother_active(N);  // step action
END_STEP
TRANSITION FROM MixDoneWaitAnother TO MixComponent
    := bContinue and not stTriblender.bComponenetMixDone;
END_TRANSITION
STEP LastComp:
    CheckIfLast_entry(P1);  // entry action
    LastComp_active(N);  // step action
    LastComp_exit(P0);  // exit action
END_STEP
TRANSITION FROM LastComp TO Init_Init_act_MixingStates
    := bContinue;
END_TRANSITION
// branch label Branch1_Init_act_MixingStates
// branch label Branch2_Init_act_MixingStates
// branch label Branch0_Init_act_MixingStates
END_ACTION

ACTION Init_Init_act_MixingStates_active:
sStateDescription	:='Triblender valve closed';
sStateInstructions	:= 'Close triblender valve';

bDisableAmount:=TRUE;
bDisableName:=TRUE;
bDisableTime:=TRUE;

wButtonColor:=16#FFC0C0C0;
stTriblender.bError:=FALSE;
stTriblender.bDisolvingDone:=FALSE;
END_ACTION

